(* CODESYS project PLC.project

Project tree, tasks and I/O mapping:
  Device : CODESYS Control Win V3 x64, CODESYS, version 3.5.20.40
    application Application
      libraries: Standard, 3.5.18.0 (System); MQTT Client Library, 3.5.20.1 (Stefan Roßmann Engineering Solutions)
      task MainTask (cyclic, interval t#20ms, priority 1) calls PLC_PRG, SCADA_PRG, PRG_MQTT
      Conveyers/
        function block Input_Conveyer [SFC]: free_entry, Create_Data
        function block Machine_Conveyer [SFC]: send_piece, recv_exit, Wait_entry, update_creation_state, recv_entry, rotate_exit, evaluate_entry, rotate_tool, process_exit, assemble_exit, swallow_entry
        function block Linear_Conveyor [SFC]: recv_entry
        function block Output_Conveyer [SFC]: Empty_Ramp, Reciving_entry, free_entry
        function block Unloading_Conveyer [SFC]: Extract_Data, wait_exit, clear_vars
        function block Loading_Conveyer [SFC]: load_entry
      program SCADA_PRG [ST]
      data type Piece
      program PLC_PRG [CFC]
      Symbols
      program AlarmManager [ST]
      global variables GVL
      program PRG_MQTT [ST]
      global variables GVL_MQTT
    Ethernet : Ethernet, CODESYS, version 4.2.0.0
      Modbus_TCP_Master : Modbus TCP Client, CODESYS, version 4.4.0.0
          settings: AutoReconnect = TRUE
        Modbus_TCP_Slave : Modbus TCP Server, CODESYS, version 4.4.0.0
            settings: Unit-ID = 255; IPAddress = [127, 0, 0, 1]; Port = 5502; InputChannel.Function Code = 2; InputChannel.Read Offset = 16#0000; InputChannel.Read Length = 140; InputChannel.Write Offset = 0; InputChannel.Write Length = 0; InputChannel.Cycle Time = 20; OutputChannel.Function Code = 15; OutputChannel.Read Offset = 0; OutputChannel.Read Length = 0; OutputChannel.Write Offset = 16#0000; OutputChannel.Write Length = 215; OutputChannel.Cycle Time = 20; pieces.Function Code = 16; pieces.Read Offset = 0; pieces.Read Length = 0; pieces.Write Offset = 16#0000; pieces.Write Length = 15; pieces.Cycle Time = 20
            input  Application.GVL.In[0] : BOOL  // InputChannel.InputChannel.Bit0
            input  Application.GVL.In[1] : BOOL  // InputChannel.InputChannel.Bit1
            input  Application.GVL.In[2] : BOOL  // InputChannel.InputChannel.Bit2
            input  Application.GVL.In[3] : BOOL  // InputChannel.InputChannel.Bit3
            input  Application.GVL.In[4] : BOOL  // InputChannel.InputChannel.Bit4
            input  Application.GVL.In[5] : BOOL  // InputChannel.InputChannel.Bit5
            input  Application.GVL.In[6] : BOOL  // InputChannel.InputChannel.Bit6
            input  Application.GVL.In[7] : BOOL  // InputChannel.InputChannel.Bit7
            input  Application.GVL.In[8] : BOOL  // InputChannel.InputChannel.Bit0
            input  Application.GVL.In[9] : BOOL  // InputChannel.InputChannel.Bit1
            input  Application.GVL.In[10] : BOOL  // InputChannel.InputChannel.Bit2
            input  Application.GVL.In[11] : BOOL  // InputChannel.InputChannel.Bit3
            input  Application.GVL.In[12] : BOOL  // InputChannel.InputChannel.Bit4
            input  Application.GVL.In[13] : BOOL  // InputChannel.InputChannel.Bit5
            input  Application.GVL.In[14] : BOOL  // InputChannel.InputChannel.Bit6
            input  Application.GVL.In[15] : BOOL  // InputChannel.InputChannel.Bit7
            input  Application.GVL.In[16] : BOOL  // InputChannel.InputChannel.Bit0
            input  Application.GVL.In[17] : BOOL  // InputChannel.InputChannel.Bit1
            input  Application.GVL.In[18] : BOOL  // InputChannel.InputChannel.Bit2
            input  Application.GVL.In[19] : BOOL  // InputChannel.InputChannel.Bit3
            input  Application.GVL.In[20] : BOOL  // InputChannel.InputChannel.Bit4
            input  Application.GVL.In[21] : BOOL  // InputChannel.InputChannel.Bit5
            input  Application.GVL.In[22] : BOOL  // InputChannel.InputChannel.Bit6
            input  Application.GVL.In[23] : BOOL  // InputChannel.InputChannel.Bit7
            input  Application.GVL.In[24] : BOOL  // InputChannel.InputChannel.Bit0
            input  Application.GVL.In[25] : BOOL  // InputChannel.InputChannel.Bit1
            input  Application.GVL.In[26] : BOOL  // InputChannel.InputChannel.Bit2
            input  Application.GVL.In[27] : BOOL  // InputChannel.InputChannel.Bit3
            input  Application.GVL.In[28] : BOOL  // InputChannel.InputChannel.Bit4
            input  Application.GVL.In[29] : BOOL  // InputChannel.InputChannel.Bit5
            input  Application.GVL.In[30] : BOOL  // InputChannel.InputChannel.Bit6
            input  Application.GVL.In[31] : BOOL  // InputChannel.InputChannel.Bit7
            input  Application.GVL.In[32] : BOOL  // InputChannel.InputChannel.Bit0
            input  Application.GVL.In[33] : BOOL  // InputChannel.InputChannel.Bit1
            input  Application.GVL.In[34] : BOOL  // InputChannel.InputChannel.Bit2
            input  Application.GVL.In[35] : BOOL  // InputChannel.InputChannel.Bit3
            input  Application.GVL.In[36] : BOOL  // InputChannel.InputChannel.Bit4
            input  Application.GVL.In[37] : BOOL  // InputChannel.InputChannel.Bit5
            input  Application.GVL.In[38] : BOOL  // InputChannel.InputChannel.Bit6
            input  Application.GVL.In[39] : BOOL  // InputChannel.InputChannel.Bit7
            input  Application.GVL.In[40] : BOOL  // InputChannel.InputChannel.Bit0
            input  Application.GVL.In[41] : BOOL  // InputChannel.InputChannel.Bit1
            input  Application.GVL.In[42] : BOOL  // InputChannel.InputChannel.Bit2
            input  Application.GVL.In[43] : BOOL  // InputChannel.InputChannel.Bit3
            input  Application.GVL.In[44] : BOOL  // InputChannel.InputChannel.Bit4
            input  Application.GVL.In[45] : BOOL  // InputChannel.InputChannel.Bit5
            input  Application.GVL.In[46] : BOOL  // InputChannel.InputChannel.Bit6
            input  Application.GVL.In[47] : BOOL  // InputChannel.InputChannel.Bit7
            input  Application.GVL.In[48] : BOOL  // InputChannel.InputChannel.Bit0
            input  Application.GVL.In[49] : BOOL  // InputChannel.InputChannel.Bit1
            input  Application.GVL.In[50] : BOOL  // InputChannel.InputChannel.Bit2
            input  Application.GVL.In[51] : BOOL  // InputChannel.InputChannel.Bit3
            input  Application.GVL.In[52] : BOOL  // InputChannel.InputChannel.Bit4
            input  Application.GVL.In[53] : BOOL  // InputChannel.InputChannel.Bit5
            input  Application.GVL.In[54] : BOOL  // InputChannel.InputChannel.Bit6
            input  Application.GVL.In[55] : BOOL  // InputChannel.InputChannel.Bit7
            input  Application.GVL.In[56] : BOOL  // InputChannel.InputChannel.Bit0
            input  Application.GVL.In[57] : BOOL  // InputChannel.InputChannel.Bit1
            input  Application.GVL.In[58] : BOOL  // InputChannel.InputChannel.Bit2
            input  Application.GVL.In[59] : BOOL  // InputChannel.InputChannel.Bit3
            input  Application.GVL.In[60] : BOOL  // InputChannel.InputChannel.Bit4
            input  Application.GVL.In[61] : BOOL  // InputChannel.InputChannel.Bit5
            input  Application.GVL.In[62] : BOOL  // InputChannel.InputChannel.Bit6
            input  Application.GVL.In[63] : BOOL  // InputChannel.InputChannel.Bit7
            input  Application.GVL.In[64] : BOOL  // InputChannel.InputChannel.Bit0
            input  Application.GVL.In[65] : BOOL  // InputChannel.InputChannel.Bit1
            input  Application.GVL.In[66] : BOOL  // InputChannel.InputChannel.Bit2
            input  Application.GVL.In[67] : BOOL  // InputChannel.InputChannel.Bit3
            input  Application.GVL.In[68] : BOOL  // InputChannel.InputChannel.Bit4
            input  Application.GVL.In[69] : BOOL  // InputChannel.InputChannel.Bit5
            input  Application.GVL.In[70] : BOOL  // InputChannel.InputChannel.Bit6
            input  Application.GVL.In[71] : BOOL  // InputChannel.InputChannel.Bit7
            input  Application.GVL.In[72] : BOOL  // InputChannel.InputChannel.Bit0
            input  Application.GVL.In[73] : BOOL  // InputChannel.InputChannel.Bit1
            input  Application.GVL.In[74] : BOOL  // InputChannel.InputChannel.Bit2
            input  Application.GVL.In[75] : BOOL  // InputChannel.InputChannel.Bit3
            input  Application.GVL.In[76] : BOOL  // InputChannel.InputChannel.Bit4
            input  Application.GVL.In[77] : BOOL  // InputChannel.InputChannel.Bit5
            input  Application.GVL.In[78] : BOOL  // InputChannel.InputChannel.Bit6
            input  Application.GVL.In[79] : BOOL  // InputChannel.InputChannel.Bit7
            input  Application.GVL.In[80] : BOOL  // InputChannel.InputChannel.Bit0
            input  Application.GVL.In[81] : BOOL  // InputChannel.InputChannel.Bit1
            input  Application.GVL.In[82] : BOOL  // InputChannel.InputChannel.Bit2
            input  Application.GVL.In[83] : BOOL  // InputChannel.InputChannel.Bit3
            input  Application.GVL.In[84] : BOOL  // InputChannel.InputChannel.Bit4
            input  Application.GVL.In[85] : BOOL  // InputChannel.InputChannel.Bit5
            input  Application.GVL.In[86] : BOOL  // InputChannel.InputChannel.Bit6
            input  Application.GVL.In[87] : BOOL  // InputChannel.InputChannel.Bit7
            input  Application.GVL.In[88] : BOOL  // InputChannel.InputChannel.Bit0
            input  Application.GVL.In[89] : BOOL  // InputChannel.InputChannel.Bit1
            input  Application.GVL.In[90] : BOOL  // InputChannel.InputChannel.Bit2
            input  Application.GVL.In[91] : BOOL  // InputChannel.InputChannel.Bit3
            input  Application.GVL.In[92] : BOOL  // InputChannel.InputChannel.Bit4
            input  Application.GVL.In[93] : BOOL  // InputChannel.InputChannel.Bit5
            input  Application.GVL.In[94] : BOOL  // InputChannel.InputChannel.Bit6
            input  Application.GVL.In[95] : BOOL  // InputChannel.InputChannel.Bit7
            input  Application.GVL.In[96] : BOOL  // InputChannel.InputChannel.Bit0
            input  Application.GVL.In[97] : BOOL  // InputChannel.InputChannel.Bit1
            input  Application.GVL.In[98] : BOOL  // InputChannel.InputChannel.Bit2
            input  Application.GVL.In[99] : BOOL  // InputChannel.InputChannel.Bit3
            input  Application.GVL.In[100] : BOOL  // InputChannel.InputChannel.Bit4
            input  Application.GVL.In[101] : BOOL  // InputChannel.InputChannel.Bit5
            input  Application.GVL.In[102] : BOOL  // InputChannel.InputChannel.Bit6
            input  Application.GVL.In[103] : BOOL  // InputChannel.InputChannel.Bit7
            input  Application.GVL.In[104] : BOOL  // InputChannel.InputChannel.Bit0
            input  Application.GVL.In[105] : BOOL  // InputChannel.InputChannel.Bit1
            input  Application.GVL.In[106] : BOOL  // InputChannel.InputChannel.Bit2
            input  Application.GVL.In[107] : BOOL  // InputChannel.InputChannel.Bit3
            input  Application.GVL.In[108] : BOOL  // InputChannel.InputChannel.Bit4
            input  Application.GVL.In[109] : BOOL  // InputChannel.InputChannel.Bit5
            input  Application.GVL.In[110] : BOOL  // InputChannel.InputChannel.Bit6
            input  Application.GVL.In[111] : BOOL  // InputChannel.InputChannel.Bit7
            input  Application.GVL.In[112] : BOOL  // InputChannel.InputChannel.Bit0
            input  Application.GVL.In[113] : BOOL  // InputChannel.InputChannel.Bit1
            input  Application.GVL.In[114] : BOOL  // InputChannel.InputChannel.Bit2
            input  Application.GVL.In[115] : BOOL  // InputChannel.InputChannel.Bit3
            input  Application.GVL.In[116] : BOOL  // InputChannel.InputChannel.Bit4
            input  Application.GVL.In[117] : BOOL  // InputChannel.InputChannel.Bit5
            input  Application.GVL.In[118] : BOOL  // InputChannel.InputChannel.Bit6
            input  Application.GVL.In[119] : BOOL  // InputChannel.InputChannel.Bit7
            input  Application.GVL.In[120] : BOOL  // InputChannel.InputChannel.Bit0
            input  Application.GVL.In[121] : BOOL  // InputChannel.InputChannel.Bit1
            input  Application.GVL.In[122] : BOOL  // InputChannel.InputChannel.Bit2
            input  Application.GVL.In[123] : BOOL  // InputChannel.InputChannel.Bit3
            input  Application.GVL.In[124] : BOOL  // InputChannel.InputChannel.Bit4
            input  Application.GVL.In[125] : BOOL  // InputChannel.InputChannel.Bit5
            input  Application.GVL.In[126] : BOOL  // InputChannel.InputChannel.Bit6
            input  Application.GVL.In[127] : BOOL  // InputChannel.InputChannel.Bit7
            input  Application.GVL.In[128] : BOOL  // InputChannel.InputChannel.Bit0
            input  Application.GVL.In[129] : BOOL  // InputChannel.InputChannel.Bit1
            input  Application.GVL.In[130] : BOOL  // InputChannel.InputChannel.Bit2
            input  Application.GVL.In[131] : BOOL  // InputChannel.InputChannel.Bit3
            input  Application.GVL.In[132] : BOOL  // InputChannel.InputChannel.Bit4
            input  Application.GVL.In[133] : BOOL  // InputChannel.InputChannel.Bit5
            input  Application.GVL.In[134] : BOOL  // InputChannel.InputChannel.Bit6
            input  Application.GVL.In[135] : BOOL  // InputChannel.InputChannel.Bit7
            input  Application.GVL.In[136] : BOOL  // InputChannel.InputChannel.Bit0
            input  Application.GVL.In[137] : BOOL  // InputChannel.InputChannel.Bit1
            input  Application.GVL.In[138] : BOOL  // InputChannel.InputChannel.Bit2
            input  Application.GVL.In[139] : BOOL  // InputChannel.InputChannel.Bit3
            output Application.GVL.Out[0] : BOOL  // OutputChannel.OutputChannel[0].Bit0
            output Application.GVL.Out[1] : BOOL  // OutputChannel.OutputChannel[0].Bit1
            output Application.GVL.Out[2] : BOOL  // OutputChannel.OutputChannel[0].Bit2
            output Application.GVL.Out[3] : BOOL  // OutputChannel.OutputChannel[0].Bit3
            output Application.GVL.Out[4] : BOOL  // OutputChannel.OutputChannel[0].Bit4
            output Application.GVL.Out[5] : BOOL  // OutputChannel.OutputChannel[0].Bit5
            output Application.GVL.Out[6] : BOOL  // OutputChannel.OutputChannel[0].Bit6
            output Application.GVL.Out[7] : BOOL  // OutputChannel.OutputChannel[0].Bit7
            output Application.GVL.Out[8] : BOOL  // OutputChannel.OutputChannel[1].Bit0
            output Application.GVL.Out[9] : BOOL  // OutputChannel.OutputChannel[1].Bit1
            output Application.GVL.Out[10] : BOOL  // OutputChannel.OutputChannel[1].Bit2
            output Application.GVL.Out[11] : BOOL  // OutputChannel.OutputChannel[1].Bit3
            output Application.GVL.Out[12] : BOOL  // OutputChannel.OutputChannel[1].Bit4
            output Application.GVL.Out[13] : BOOL  // OutputChannel.OutputChannel[1].Bit5
            output Application.GVL.Out[14] : BOOL  // OutputChannel.OutputChannel[1].Bit6
            output Application.GVL.Out[15] : BOOL  // OutputChannel.OutputChannel[1].Bit7
            output Application.GVL.Out[16] : BOOL  // OutputChannel.OutputChannel[2].Bit0
            output Application.GVL.Out[17] : BOOL  // OutputChannel.OutputChannel[2].Bit1
            output Application.GVL.Out[18] : BOOL  // OutputChannel.OutputChannel[2].Bit2
            output Application.GVL.Out[19] : BOOL  // OutputChannel.OutputChannel[2].Bit3
            output Application.GVL.Out[20] : BOOL  // OutputChannel.OutputChannel[2].Bit4
            output Application.GVL.Out[21] : BOOL  // OutputChannel.OutputChannel[2].Bit5
            output Application.GVL.Out[22] : BOOL  // OutputChannel.OutputChannel[2].Bit6
            output Application.GVL.Out[23] : BOOL  // OutputChannel.OutputChannel[2].Bit7
            output Application.GVL.Out[24] : BOOL  // OutputChannel.OutputChannel[3].Bit0
            output Application.GVL.Out[25] : BOOL  // OutputChannel.OutputChannel[3].Bit1
            output Application.GVL.Out[26] : BOOL  // OutputChannel.OutputChannel[3].Bit2
            output Application.GVL.Out[27] : BOOL  // OutputChannel.OutputChannel[3].Bit3
            output Application.GVL.Out[28] : BOOL  // OutputChannel.OutputChannel[3].Bit4
            output Application.GVL.Out[29] : BOOL  // OutputChannel.OutputChannel[3].Bit5
            output Application.GVL.Out[30] : BOOL  // OutputChannel.OutputChannel[3].Bit6
            output Application.GVL.Out[31] : BOOL  // OutputChannel.OutputChannel[3].Bit7
            output Application.GVL.Out[32] : BOOL  // OutputChannel.OutputChannel[4].Bit0
            output Application.GVL.Out[33] : BOOL  // OutputChannel.OutputChannel[4].Bit1
            output Application.GVL.Out[34] : BOOL  // OutputChannel.OutputChannel[4].Bit2
            output Application.GVL.Out[35] : BOOL  // OutputChannel.OutputChannel[4].Bit3
            output Application.GVL.Out[36] : BOOL  // OutputChannel.OutputChannel[4].Bit4
            output Application.GVL.Out[37] : BOOL  // OutputChannel.OutputChannel[4].Bit5
            output Application.GVL.Out[38] : BOOL  // OutputChannel.OutputChannel[4].Bit6
            output Application.GVL.Out[39] : BOOL  // OutputChannel.OutputChannel[4].Bit7
            output Application.GVL.Out[40] : BOOL  // OutputChannel.OutputChannel[5].Bit0
            output Application.GVL.Out[41] : BOOL  // OutputChannel.OutputChannel[5].Bit1
            output Application.GVL.Out[42] : BOOL  // OutputChannel.OutputChannel[5].Bit2
            output Application.GVL.Out[43] : BOOL  // OutputChannel.OutputChannel[5].Bit3
            output Application.GVL.Out[44] : BOOL  // OutputChannel.OutputChannel[5].Bit4
            output Application.GVL.Out[45] : BOOL  // OutputChannel.OutputChannel[5].Bit5
            output Application.GVL.Out[46] : BOOL  // OutputChannel.OutputChannel[5].Bit6
            output Application.GVL.Out[47] : BOOL  // OutputChannel.OutputChannel[5].Bit7
            output Application.GVL.Out[48] : BOOL  // OutputChannel.OutputChannel[6].Bit0
            output Application.GVL.Out[49] : BOOL  // OutputChannel.OutputChannel[6].Bit1
            output Application.GVL.Out[50] : BOOL  // OutputChannel.OutputChannel[6].Bit2
            output Application.GVL.Out[51] : BOOL  // OutputChannel.OutputChannel[6].Bit3
            output Application.GVL.Out[52] : BOOL  // OutputChannel.OutputChannel[6].Bit4
            output Application.GVL.Out[53] : BOOL  // OutputChannel.OutputChannel[6].Bit5
            output Application.GVL.Out[54] : BOOL  // OutputChannel.OutputChannel[6].Bit6
            output Application.GVL.Out[55] : BOOL  // OutputChannel.OutputChannel[6].Bit7
            output Application.GVL.Out[56] : BOOL  // OutputChannel.OutputChannel[7].Bit0
            output Application.GVL.Out[57] : BOOL  // OutputChannel.OutputChannel[7].Bit1
            output Application.GVL.Out[58] : BOOL  // OutputChannel.OutputChannel[7].Bit2
            output Application.GVL.Out[59] : BOOL  // OutputChannel.OutputChannel[7].Bit3
            output Application.GVL.Out[60] : BOOL  // OutputChannel.OutputChannel[7].Bit4
            output Application.GVL.Out[61] : BOOL  // OutputChannel.OutputChannel[7].Bit5
            output Application.GVL.Out[62] : BOOL  // OutputChannel.OutputChannel[7].Bit6
            output Application.GVL.Out[63] : BOOL  // OutputChannel.OutputChannel[7].Bit7
            output Application.GVL.Out[64] : BOOL  // OutputChannel.OutputChannel[8].Bit0
            output Application.GVL.Out[65] : BOOL  // OutputChannel.OutputChannel[8].Bit1
            output Application.GVL.Out[66] : BOOL  // OutputChannel.OutputChannel[8].Bit2
            output Application.GVL.Out[67] : BOOL  // OutputChannel.OutputChannel[8].Bit3
            output Application.GVL.Out[68] : BOOL  // OutputChannel.OutputChannel[8].Bit4
            output Application.GVL.Out[69] : BOOL  // OutputChannel.OutputChannel[8].Bit5
            output Application.GVL.Out[70] : BOOL  // OutputChannel.OutputChannel[8].Bit6
            output Application.GVL.Out[71] : BOOL  // OutputChannel.OutputChannel[8].Bit7
            output Application.GVL.Out[72] : BOOL  // OutputChannel.OutputChannel[9].Bit0
            output Application.GVL.Out[73] : BOOL  // OutputChannel.OutputChannel[9].Bit1
            output Application.GVL.Out[74] : BOOL  // OutputChannel.OutputChannel[9].Bit2
            output Application.GVL.Out[75] : BOOL  // OutputChannel.OutputChannel[9].Bit3
            output Application.GVL.Out[76] : BOOL  // OutputChannel.OutputChannel[9].Bit4
            output Application.GVL.Out[77] : BOOL  // OutputChannel.OutputChannel[9].Bit5
            output Application.GVL.Out[78] : BOOL  // OutputChannel.OutputChannel[9].Bit6
            output Application.GVL.Out[79] : BOOL  // OutputChannel.OutputChannel[9].Bit7
            output Application.GVL.Out[80] : BOOL  // OutputChannel.OutputChannel[10].Bit0
            output Application.GVL.Out[81] : BOOL  // OutputChannel.OutputChannel[10].Bit1
            output Application.GVL.Out[82] : BOOL  // OutputChannel.OutputChannel[10].Bit2
            output Application.GVL.Out[83] : BOOL  // OutputChannel.OutputChannel[10].Bit3
            output Application.GVL.Out[84] : BOOL  // OutputChannel.OutputChannel[10].Bit4
            output Application.GVL.Out[85] : BOOL  // OutputChannel.OutputChannel[10].Bit5
            output Application.GVL.Out[86] : BOOL  // OutputChannel.OutputChannel[10].Bit6
            output Application.GVL.Out[87] : BOOL  // OutputChannel.OutputChannel[10].Bit7
            output Application.GVL.Out[88] : BOOL  // OutputChannel.OutputChannel[11].Bit0
            output Application.GVL.Out[89] : BOOL  // OutputChannel.OutputChannel[11].Bit1
            output Application.GVL.Out[90] : BOOL  // OutputChannel.OutputChannel[11].Bit2
            output Application.GVL.Out[91] : BOOL  // OutputChannel.OutputChannel[11].Bit3
            output Application.GVL.Out[92] : BOOL  // OutputChannel.OutputChannel[11].Bit4
            output Application.GVL.Out[93] : BOOL  // OutputChannel.OutputChannel[11].Bit5
            output Application.GVL.Out[94] : BOOL  // OutputChannel.OutputChannel[11].Bit6
            output Application.GVL.Out[95] : BOOL  // OutputChannel.OutputChannel[11].Bit7
            output Application.GVL.Out[96] : BOOL  // OutputChannel.OutputChannel[12].Bit0
            output Application.GVL.Out[97] : BOOL  // OutputChannel.OutputChannel[12].Bit1
            output Application.GVL.Out[98] : BOOL  // OutputChannel.OutputChannel[12].Bit2
            output Application.GVL.Out[99] : BOOL  // OutputChannel.OutputChannel[12].Bit3
            output Application.GVL.Out[100] : BOOL  // OutputChannel.OutputChannel[12].Bit4
            output Application.GVL.Out[101] : BOOL  // OutputChannel.OutputChannel[12].Bit5
            output Application.GVL.Out[102] : BOOL  // OutputChannel.OutputChannel[12].Bit6
            output Application.GVL.Out[103] : BOOL  // OutputChannel.OutputChannel[12].Bit7
            output Application.GVL.Out[104] : BOOL  // OutputChannel.OutputChannel[13].Bit0
            output Application.GVL.Out[105] : BOOL  // OutputChannel.OutputChannel[13].Bit1
            output Application.GVL.Out[106] : BOOL  // OutputChannel.OutputChannel[13].Bit2
            output Application.GVL.Out[107] : BOOL  // OutputChannel.OutputChannel[13].Bit3
            output Application.GVL.Out[108] : BOOL  // OutputChannel.OutputChannel[13].Bit4
            output Application.GVL.Out[109] : BOOL  // OutputChannel.OutputChannel[13].Bit5
            output Application.GVL.Out[110] : BOOL  // OutputChannel.OutputChannel[13].Bit6
            output Application.GVL.Out[111] : BOOL  // OutputChannel.OutputChannel[13].Bit7
            output Application.GVL.Out[112] : BOOL  // OutputChannel.OutputChannel[14].Bit0
            output Application.GVL.Out[113] : BOOL  // OutputChannel.OutputChannel[14].Bit1
            output Application.GVL.Out[114] : BOOL  // OutputChannel.OutputChannel[14].Bit2
            output Application.GVL.Out[115] : BOOL  // OutputChannel.OutputChannel[14].Bit3
            output Application.GVL.Out[116] : BOOL  // OutputChannel.OutputChannel[14].Bit4
            output Application.GVL.Out[117] : BOOL  // OutputChannel.OutputChannel[14].Bit5
            output Application.GVL.Out[118] : BOOL  // OutputChannel.OutputChannel[14].Bit6
            output Application.GVL.Out[119] : BOOL  // OutputChannel.OutputChannel[14].Bit7
            output Application.GVL.Out[120] : BOOL  // OutputChannel.OutputChannel[15].Bit0
            output Application.GVL.Out[121] : BOOL  // OutputChannel.OutputChannel[15].Bit1
            output Application.GVL.Out[122] : BOOL  // OutputChannel.OutputChannel[15].Bit2
            output Application.GVL.Out[123] : BOOL  // OutputChannel.OutputChannel[15].Bit3
            output Application.GVL.Out[124] : BOOL  // OutputChannel.OutputChannel[15].Bit4
            output Application.GVL.Out[125] : BOOL  // OutputChannel.OutputChannel[15].Bit5
            output Application.GVL.Out[126] : BOOL  // OutputChannel.OutputChannel[15].Bit6
            output Application.GVL.Out[127] : BOOL  // OutputChannel.OutputChannel[15].Bit7
            output Application.GVL.Out[128] : BOOL  // OutputChannel.OutputChannel[16].Bit0
            output Application.GVL.Out[129] : BOOL  // OutputChannel.OutputChannel[16].Bit1
            output Application.GVL.Out[130] : BOOL  // OutputChannel.OutputChannel[16].Bit2
            output Application.GVL.Out[131] : BOOL  // OutputChannel.OutputChannel[16].Bit3
            output Application.GVL.Out[132] : BOOL  // OutputChannel.OutputChannel[16].Bit4
            output Application.GVL.Out[133] : BOOL  // OutputChannel.OutputChannel[16].Bit5
            output Application.GVL.Out[134] : BOOL  // OutputChannel.OutputChannel[16].Bit6
            output Application.GVL.Out[135] : BOOL  // OutputChannel.OutputChannel[16].Bit7
            output Application.GVL.Out[136] : BOOL  // OutputChannel.OutputChannel[17].Bit0
            output Application.GVL.Out[137] : BOOL  // OutputChannel.OutputChannel[17].Bit1
            output Application.GVL.Out[138] : BOOL  // OutputChannel.OutputChannel[17].Bit2
            output Application.GVL.Out[139] : BOOL  // OutputChannel.OutputChannel[17].Bit3
            output Application.GVL.Out[140] : BOOL  // OutputChannel.OutputChannel[17].Bit4
            output Application.GVL.Out[141] : BOOL  // OutputChannel.OutputChannel[17].Bit5
            output Application.GVL.Out[142] : BOOL  // OutputChannel.OutputChannel[17].Bit6
            output Application.GVL.Out[143] : BOOL  // OutputChannel.OutputChannel[17].Bit7
            output Application.GVL.Out[144] : BOOL  // OutputChannel.OutputChannel[18].Bit0
            output Application.GVL.Out[145] : BOOL  // OutputChannel.OutputChannel[18].Bit1
            output Application.GVL.Out[146] : BOOL  // OutputChannel.OutputChannel[18].Bit2
            output Application.GVL.Out[147] : BOOL  // OutputChannel.OutputChannel[18].Bit3
            output Application.GVL.Out[148] : BOOL  // OutputChannel.OutputChannel[18].Bit4
            output Application.GVL.Out[149] : BOOL  // OutputChannel.OutputChannel[18].Bit5
            output Application.GVL.Out[150] : BOOL  // OutputChannel.OutputChannel[18].Bit6
            output Application.GVL.Out[151] : BOOL  // OutputChannel.OutputChannel[18].Bit7
            output Application.GVL.Out[152] : BOOL  // OutputChannel.OutputChannel[19].Bit0
            output Application.GVL.Out[153] : BOOL  // OutputChannel.OutputChannel[19].Bit1
            output Application.GVL.Out[154] : BOOL  // OutputChannel.OutputChannel[19].Bit2
            output Application.GVL.Out[155] : BOOL  // OutputChannel.OutputChannel[19].Bit3
            output Application.GVL.Out[156] : BOOL  // OutputChannel.OutputChannel[19].Bit4
            output Application.GVL.Out[157] : BOOL  // OutputChannel.OutputChannel[19].Bit5
            output Application.GVL.Out[158] : BOOL  // OutputChannel.OutputChannel[19].Bit6
            output Application.GVL.Out[159] : BOOL  // OutputChannel.OutputChannel[19].Bit7
            output Application.GVL.Out[160] : BOOL  // OutputChannel.OutputChannel[20].Bit0
            output Application.GVL.Out[161] : BOOL  // OutputChannel.OutputChannel[20].Bit1
            output Application.GVL.Out[162] : BOOL  // OutputChannel.OutputChannel[20].Bit2
            output Application.GVL.Out[163] : BOOL  // OutputChannel.OutputChannel[20].Bit3
            output Application.GVL.Out[164] : BOOL  // OutputChannel.OutputChannel[20].Bit4
            output Application.GVL.Out[165] : BOOL  // OutputChannel.OutputChannel[20].Bit5
            output Application.GVL.Out[166] : BOOL  // OutputChannel.OutputChannel[20].Bit6
            output Application.GVL.Out[167] : BOOL  // OutputChannel.OutputChannel[20].Bit7
            output Application.GVL.Out[168] : BOOL  // OutputChannel.OutputChannel[21].Bit0
            output Application.GVL.Out[169] : BOOL  // OutputChannel.OutputChannel[21].Bit1
            output Application.GVL.Out[170] : BOOL  // OutputChannel.OutputChannel[21].Bit2
            output Application.GVL.Out[171] : BOOL  // OutputChannel.OutputChannel[21].Bit3
            output Application.GVL.Out[172] : BOOL  // OutputChannel.OutputChannel[21].Bit4
            output Application.GVL.Out[173] : BOOL  // OutputChannel.OutputChannel[21].Bit5
            output Application.GVL.Out[174] : BOOL  // OutputChannel.OutputChannel[21].Bit6
            output Application.GVL.Out[175] : BOOL  // OutputChannel.OutputChannel[21].Bit7
            output Application.GVL.Out[176] : BOOL  // OutputChannel.OutputChannel[22].Bit0
            output Application.GVL.Out[177] : BOOL  // OutputChannel.OutputChannel[22].Bit1
            output Application.GVL.Out[178] : BOOL  // OutputChannel.OutputChannel[22].Bit2
            output Application.GVL.Out[179] : BOOL  // OutputChannel.OutputChannel[22].Bit3
            output Application.GVL.Out[180] : BOOL  // OutputChannel.OutputChannel[22].Bit4
            output Application.GVL.Out[181] : BOOL  // OutputChannel.OutputChannel[22].Bit5
            output Application.GVL.Out[182] : BOOL  // OutputChannel.OutputChannel[22].Bit6
            output Application.GVL.Out[183] : BOOL  // OutputChannel.OutputChannel[22].Bit7
            output Application.GVL.Out[184] : BOOL  // OutputChannel.OutputChannel[23].Bit0
            output Application.GVL.Out[185] : BOOL  // OutputChannel.OutputChannel[23].Bit1
            output Application.GVL.Out[186] : BOOL  // OutputChannel.OutputChannel[23].Bit2
            output Application.GVL.Out[187] : BOOL  // OutputChannel.OutputChannel[23].Bit3
            output Application.GVL.Out[188] : BOOL  // OutputChannel.OutputChannel[23].Bit4
            output Application.GVL.Out[189] : BOOL  // OutputChannel.OutputChannel[23].Bit5
            output Application.GVL.Out[190] : BOOL  // OutputChannel.OutputChannel[23].Bit6
            output Application.GVL.Out[191] : BOOL  // OutputChannel.OutputChannel[23].Bit7
            output Application.GVL.Out[192] : BOOL  // OutputChannel.OutputChannel[24].Bit0
            output Application.GVL.Out[193] : BOOL  // OutputChannel.OutputChannel[24].Bit1
            output Application.GVL.Out[194] : BOOL  // OutputChannel.OutputChannel[24].Bit2
            output Application.GVL.Out[195] : BOOL  // OutputChannel.OutputChannel[24].Bit3
            output Application.GVL.Out[196] : BOOL  // OutputChannel.OutputChannel[24].Bit4
            output Application.GVL.Out[197] : BOOL  // OutputChannel.OutputChannel[24].Bit5
            output Application.GVL.Out[198] : BOOL  // OutputChannel.OutputChannel[24].Bit6
            output Application.GVL.Out[199] : BOOL  // OutputChannel.OutputChannel[24].Bit7
            output Application.GVL.Out[200] : BOOL  // OutputChannel.OutputChannel[25].Bit0
            output Application.GVL.Out[201] : BOOL  // OutputChannel.OutputChannel[25].Bit1
            output Application.GVL.Out[202] : BOOL  // OutputChannel.OutputChannel[25].Bit2
            output Application.GVL.Out[203] : BOOL  // OutputChannel.OutputChannel[25].Bit3
            output Application.GVL.Out[204] : BOOL  // OutputChannel.OutputChannel[25].Bit4
            output Application.GVL.Out[205] : BOOL  // OutputChannel.OutputChannel[25].Bit5
            output Application.GVL.Out[206] : BOOL  // OutputChannel.OutputChannel[25].Bit6
            output Application.GVL.Out[207] : BOOL  // OutputChannel.OutputChannel[25].Bit7
            output Application.GVL.Out[208] : BOOL  // OutputChannel.OutputChannel[26].Bit0
            output Application.GVL.Out[209] : BOOL  // OutputChannel.OutputChannel[26].Bit1
            output Application.GVL.Out[210] : BOOL  // OutputChannel.OutputChannel[26].Bit2
            output Application.GVL.Out[211] : BOOL  // OutputChannel.OutputChannel[26].Bit3
            output Application.GVL.Out[212] : BOOL  // OutputChannel.OutputChannel[26].Bit4
            output Application.GVL.Out[213] : BOOL  // OutputChannel.OutputChannel[26].Bit5
            output Application.GVL.Out[214] : BOOL  // OutputChannel.OutputChannel[26].Bit6
            output Application.GVL.Reg[0] : WORD  // pieces.pieces[0]
            output Application.GVL.Reg[1] : WORD  // pieces.pieces[1]
            output Application.GVL.Reg[2] : WORD  // pieces.pieces[2]
            output Application.GVL.Reg[3] : WORD  // pieces.pieces[3]
            output Application.GVL.Reg[4] : WORD  // pieces.pieces[4]
            output Application.GVL.Reg[5] : WORD  // pieces.pieces[5]
            output Application.GVL.Reg[6] : WORD  // pieces.pieces[6]
            output Application.GVL.Reg[7] : WORD  // pieces.pieces[7]
            output Application.GVL.Reg[8] : WORD  // pieces.pieces[8]
            output Application.GVL.Reg[9] : WORD  // pieces.pieces[9]
            output Application.GVL.Reg[10] : WORD  // pieces.pieces[10]
            output Application.GVL.Reg[11] : WORD  // pieces.pieces[11]
            output Application.GVL.Reg[12] : WORD  // pieces.pieces[12]
            output Application.GVL.Reg[13] : WORD  // pieces.pieces[13]
            output Application.GVL.Reg[14] : WORD  // pieces.pieces[14]
            unmapped channels: InputChannel, OutputChannel, pieces
      ModbusTCP_Slave_Device : ModbusTCP Server Device, CODESYS, version 4.4.0.0
          settings: UpdateableHolding = TRUE; DistinctBitAreas = TRUE; Coils Size = 48; Discrete Inputs Size = 8
          output S_sensor1 : BOOL  // Holding Registers.Holding Registers.Bit0
          output S_sensor2 : BOOL  // Holding Registers.Holding Registers.Bit1
          output S_sensor3 : BOOL  // Holding Registers.Holding Registers.Bit2
          output C1_stop : BOOL  // Holding Registers.Holding Registers.Bit0
          output C2_stop : BOOL  // Holding Registers.Holding Registers.Bit1
          output C3_stop : BOOL  // Holding Registers.Holding Registers.Bit2
          output In_on : BOOL  // Coils.Coils.Bit0
          output M1a_on : BOOL  // Coils.Coils.Bit1
          output L1_on : BOOL  // Coils.Coils.Bit2
          output M1b_on : BOOL  // Coils.Coils.Bit3
          output L2_on : BOOL  // Coils.Coils.Bit4
          output M1c_on : BOOL  // Coils.Coils.Bit5
          output Out_on : BOOL  // Coils.Coils.Bit6
          output C1_In_Sensor : BOOL  // Coils.Coils.Bit7
          output M1a_Sensor : BOOL  // Coils.Coils.Bit0
          output C1_L1_Sensor : BOOL  // Coils.Coils.Bit1
          output M1b_Sensor : BOOL  // Coils.Coils.Bit2
          output C1_L2_Sensor : BOOL  // Coils.Coils.Bit3
          output M1c_Sensor : BOOL  // Coils.Coils.Bit4
          output M1a_T1 : BOOL  // Coils.Coils.Bit5
          output M1a_T2 : BOOL  // Coils.Coils.Bit6
          output M1a_T3 : BOOL  // Coils.Coils.Bit7
          output C1_Out_Sensor : BOOL  // Coils.Coils.Bit0
          output M1a_done : BOOL  // Coils.Coils.Bit1
          output M1a_Idle_Alarm : BOOL  // Coils.Coils.Bit2
          output M1a_Manual : BOOL  // Coils.Coils.Bit3
          output M1a_Auto : BOOL  // Coils.Coils.Bit4
          output M1c_T11 : BOOL  // Coils.Coils.Bit5
          output M1a_Manutencao : BOOL  // Coils.Coils.Bit6
          unmapped channels: Holding Registers, Input Registers, Coils, Discrete Inputs
*)

// Device/Application/Piece
TYPE Piece :
STRUCT
	/// 0=Empty, 1=Wood, 2=Metal, 3=RtopW, 4=STopW, 5=LegW, 6=RtopM, 7=STopM, 8=LegM, 9=RWW, 10=SWW, 11=RWM, 12=SWM, 13=RMM, 14=SMM
	Type_ID: UINT;
	/// TRUE if piece is destroyed 
	Is_Black: BOOL;
END_STRUCT
END_TYPE

// Device/Application/GVL
VAR_GLOBAL
	In: ARRAY[0..139] OF BOOL;
	Out: ARRAY[0..220] OF BOOL;
	Reg: ARRAY[0..15] OF UINT;
	WareHouseTop: ARRAY[0..31] OF Piece;
	WareHouseBottom: ARRAY[0..31] OF Piece;
	/// Number of pieces currently in W1
	W1_Count: UINT := 0;
	/// Number of pieces currently in W2~
	W2_Count: UINT := 0;
	
	Tool_M1a: ARRAY[0..2] OF INT := [1, 2, 3];
	Tool_Time: ARRAY[0..11] OF TIME := [T#0S, T#30S, T#20S, T#10S, T#35S, T#30S, T#25S, T#0S, T#10S, T#10S, T#30S, T#40S];
	Tool_M1b: ARRAY[0..2] OF INT := [1, 2, 3];
	Tool_M1c: ARRAY[0..2] OF INT := [8, 9, 11];
	Tool_M2a: ARRAY[0..2] OF INT := [1, 2, 3];
	Tool_M2b: ARRAY[0..2] OF INT := [1, 2, 3];
	Tool_M2c: ARRAY[0..2] OF INT := [8, 9, 10];
	Tool_M3a: ARRAY[0..2] OF INT := [4, 5, 6];
	Tool_M3b: ARRAY[0..2] OF INT := [4, 5, 6];
	Tool_M3c: ARRAY[0..2] OF INT := [8, 9, 11];
	Tool_M4a: ARRAY[0..2] OF INT := [4, 5, 6];
	Tool_M4b: ARRAY[0..2] OF INT := [4, 5, 6];
	Tool_M4c: ARRAY[0..2] OF INT := [8, 9, 10];
END_VAR

// Device/Application/GVL_MQTT
(*
  GVL_MQTT — Global Variable List for ThingsBoard MQTT connection
  Paste this into a new GVL named "GVL_MQTT" in CODESYS.
  Requires: MQTT Client Library (namespace: MQTT_Client) in Library Manager.
*)

VAR_GLOBAL
    // Publisher — sends PLC I/O telemetry to ThingsBoard PLC_Gateway device
    fbMQTT_Pub          : MQTT_Client.FB_MQTTClient;

    // Subscriber — receives RPC commands from ThingsBoard
    fbMQTT_Sub          : MQTT_Client.FB_MQTTClient;

    // 2-second publish timer
    tPublishTimer       : TON;

    // Publish group counter (1=inputs, 2=unload req, 3=unload type, 4=warehouse)
    nPublishGroup       : INT := 0;

    // RPC command handling
    sRPCMessage         : STRING(1024);
    bNewRPC             : BOOL;
	
END_VAR

// Device/Application/PLC_PRG
PROGRAM PLC_PRG
VAR
	C1: Linear_Conveyor;
	C2: Linear_Conveyor;
	C3: Linear_Conveyor;
	C4: Linear_Conveyor;
	C5: Linear_Conveyor;
	C7: Linear_Conveyor;
	C9: Linear_Conveyor;
	C12: Linear_Conveyor;
	C14: Linear_Conveyor;
	C17: Linear_Conveyor;
	C19: Linear_Conveyor;
	C22: Linear_Conveyor;
	C24: Linear_Conveyor;
	C6: Machine_Conveyer;
	C8: Machine_Conveyer;
	C10: Machine_Conveyer;
	C11: Machine_Conveyer;
	C13: Machine_Conveyer;
	C15: Machine_Conveyer;
	C16: Machine_Conveyer;
	C18: Machine_Conveyer;
	C20: Machine_Conveyer;
	C21: Machine_Conveyer;
	C23: Machine_Conveyer;
	C25: Machine_Conveyer;
	O1: Output_Conveyer;
	O2: Output_Conveyer;
	O3: Output_Conveyer;
	O4: Output_Conveyer;
	O5: Output_Conveyer;
	I1: Input_Conveyer;
	I2: Input_Conveyer;
	I3: Input_Conveyer;
	I4: Input_Conveyer;
	I5: Input_Conveyer;
	U1: Unloading_Conveyer;
	U2: Unloading_Conveyer;
	U3: Unloading_Conveyer;
	U4: Unloading_Conveyer;
	U5: Unloading_Conveyer;
	U6: Unloading_Conveyer;
	U7: Unloading_Conveyer;
	U8: Unloading_Conveyer;
	U9: Unloading_Conveyer;
	U10: Unloading_Conveyer;
	L1: Loading_Conveyer;
	L2: Loading_Conveyer;
	L3: Loading_Conveyer;
	L4: Loading_Conveyer;
	L5: Loading_Conveyer;
	L6: Loading_Conveyer;
	L7: Loading_Conveyer;
	L8: Loading_Conveyer;
	L9: Loading_Conveyer;
	L10: Loading_Conveyer;
	piece_material_I1: UINT;
	piece_material_I2: UINT;
	piece_material_I3: UINT;
	piece_material_I4: UINT;
	piece_material_I5: UINT;
	piece_material_U1: UINT;
	piece_material_U2: UINT;
	piece_material_U3: UINT;
	piece_material_U4: UINT;
	piece_material_U5: UINT;
	piece_material_U6: UINT;
	piece_material_U7: UINT;
	piece_material_U8: UINT;
	piece_material_U9: UINT;
	piece_material_U10: UINT;
	Create_Piece_I1: BOOL;
	Create_Piece_I2: BOOL;
	Create_Piece_I3: BOOL;
	Create_Piece_I4: BOOL;
	Create_Piece_I5: BOOL;
	Unload_Req_U1: BOOL;
	Unload_Req_U2: BOOL;
	Unload_Req_U3: BOOL;
	Unload_Req_U4: BOOL;
	Unload_Req_U5: BOOL;
	Unload_Req_U6: BOOL;
	Unload_Req_U7: BOOL;
	Unload_Req_U8: BOOL;
	Unload_Req_U9: BOOL;
	Unload_Req_U10: BOOL;
	Unload_Type_U1: UINT;
	Unload_Type_U2: UINT;
	Unload_Type_U3: UINT;
	Unload_Type_U4: UINT;
	Unload_Type_U5: UINT;
	Unload_Type_U6: UINT;
	Unload_Type_U7: UINT;
	Unload_Type_U8: UINT;
	Unload_Type_U9: UINT;
	Unload_Type_U10: UINT;
	Output_Unload_O1: BOOL;
	Output_Unload_O2: BOOL;
	Output_Unload_O3: BOOL;
	Output_Unload_O4: BOOL;
	Output_Unload_O5: BOOL;
END_VAR

I1(
    Ioff := 0,
    Qoff := 0,
    Create_Piece := Create_Piece_I1,
    piece_material := piece_material_I1,
    free_I := L6.free_O,
    reg_numb := 0); // Input_Conveyer
L6(Ioff := 5, Qoff := 10, Target_WH := 1, Direction := 1, Piece_In := I1.Piece_Out, recv_I := I1.recv_O); // Loading_Conveyer
I2(
    Ioff := 1,
    Qoff := 2,
    Create_Piece := Create_Piece_I2,
    piece_material := piece_material_I2,
    free_I := L7.free_O,
    reg_numb := 1); // Input_Conveyer
L7(Ioff := 6, Qoff := 13, Target_WH := 1, Direction := 1, Piece_In := I2.Piece_Out, recv_I := I2.recv_O); // Loading_Conveyer
I3(
    Ioff := 2,
    Qoff := 4,
    Create_Piece := Create_Piece_I3,
    piece_material := piece_material_I3,
    free_I := L8.free_O,
    reg_numb := 2); // Input_Conveyer
L8(Ioff := 7, Qoff := 16, Target_WH := 1, Direction := 1, Piece_In := I3.Piece_Out, recv_I := I3.recv_O); // Loading_Conveyer
I4(
    Ioff := 3,
    Qoff := 6,
    Create_Piece := Create_Piece_I4,
    piece_material := piece_material_I4,
    free_I := L9.free_O,
    reg_numb := 3); // Input_Conveyer
L9(Ioff := 8, Qoff := 19, Target_WH := 1, Direction := 1, Piece_In := I4.Piece_Out, recv_I := I4.recv_O); // Loading_Conveyer
I5(
    Ioff := 4,
    Qoff := 8,
    Create_Piece := Create_Piece_I5,
    piece_material := piece_material_I5,
    free_I := L10.free_O,
    reg_numb := 4); // Input_Conveyer
L10(Ioff := 9, Qoff := 22, Target_WH := 1, Direction := 1, Piece_In := I5.Piece_Out, recv_I := I5.recv_O); // Loading_Conveyer
L1(Ioff := 10, Qoff := 25, Target_WH := 1, Direction := 0, Piece_In := C1.Passed_Piece, recv_I := C1.recv_O); // Loading_Conveyer
U2(
    Ioff := 11,
    Qoff := 28,
    Target_WH := 1,
    Direction := 1,
    Unload_Req := Unload_Req_U2,
    free_I := C6.free_O,
    piece_material := Unload_Type_U2,
    reg_numb := 5); // Unloading_Conveyer
U3(
    Ioff := 12,
    Qoff := 30,
    Target_WH := 1,
    Direction := 1,
    Unload_Req := Unload_Req_U3,
    free_I := C11.free_O,
    piece_material := Unload_Type_U3,
    reg_numb := 6); // Unloading_Conveyer
U4(
    Ioff := 13,
    Qoff := 32,
    Target_WH := 1,
    Direction := 1,
    Unload_Req := Unload_Req_U4,
    free_I := C16.free_O,
    piece_material := Unload_Type_U4,
    reg_numb := 7); // Unloading_Conveyer
U5(
    Ioff := 14,
    Qoff := 34,
    Target_WH := 1,
    Direction := 1,
    Unload_Req := Unload_Req_U5,
    free_I := C21.free_O,
    piece_material := Unload_Type_U5,
    reg_numb := 8); // Unloading_Conveyer
C1(
    Ioff := 25,
    Qoff := 60,
    Direction := 0,
    Piece_Type := C2.Passed_Piece,
    recv_I := C2.recv_O,
    free_I := L1.free_O); // Linear_Conveyor
C6(
    Ioff := 30,
    Qoff := 70,
    Piece_In := U2.Piece_Out,
    recv_I := U2.recv_O,
    Direction := 1,
    free_I := C7.free_O,
    Tool_Magazine := GVL.Tool_M1a); // Machine_Conveyer
C11(
    Ioff := 50,
    Qoff := 104,
    Piece_In := U3.Piece_Out,
    recv_I := U3.recv_O,
    Direction := 1,
    free_I := C12.free_O,
    Tool_Magazine := GVL.Tool_M2a); // Machine_Conveyer
C16(
    Ioff := 70,
    Qoff := 138,
    Piece_In := U4.Piece_Out,
    recv_I := U4.recv_O,
    Direction := 1,
    free_I := C17.free_O,
    Tool_Magazine := GVL.Tool_M3a); // Machine_Conveyer
C21(
    Ioff := 90,
    Qoff := 172,
    Piece_In := U5.Piece_Out,
    Direction := 1,
    recv_I := U5.recv_O,
    free_I := C22.free_O,
    Tool_Magazine := GVL.Tool_M4a); // Machine_Conveyer
C2(
    Ioff := 26,
    Qoff := 62,
    Direction := 0,
    Piece_Type := C3.Passed_Piece,
    recv_I := C3.recv_O,
    free_I := C1.free_O); // Linear_Conveyor
C7(
    Ioff := 36,
    Qoff := 80,
    Direction := 1,
    Piece_Type := C6.Piece_Out,
    recv_I := C6.recv_O,
    free_I := C8.free_O); // Linear_Conveyor
C12(
    Ioff := 56,
    Qoff := 114,
    Direction := 1,
    Piece_Type := C11.Piece_Out,
    recv_I := C11.recv_O,
    free_I := C13.free_O); // Linear_Conveyor
C17(
    Ioff := 76,
    Qoff := 148,
    Direction := 1,
    Piece_Type := C16.Piece_Out,
    recv_I := C16.recv_O,
    free_I := C18.free_O); // Linear_Conveyor
C22(
    Ioff := 96,
    Qoff := 182,
    Direction := 1,
    Piece_Type := C21.Piece_Out,
    recv_I := C21.recv_O,
    free_I := C23.free_O); // Linear_Conveyor
C3(
    Ioff := 27,
    Qoff := 64,
    Direction := 0,
    Piece_Type := C4.Passed_Piece,
    recv_I := C4.recv_O,
    free_I := C2.free_O); // Linear_Conveyor
C8(
    Ioff := 37,
    Qoff := 82,
    Piece_In := C7.Passed_Piece,
    Direction := 1,
    recv_I := C7.recv_O,
    free_I := C9.free_O,
    Tool_Magazine := GVL.Tool_M1b); // Machine_Conveyer
C13(
    Ioff := 57,
    Qoff := 116,
    Piece_In := C12.Passed_Piece,
    Direction := 1,
    recv_I := C12.recv_O,
    free_I := C14.free_O,
    Tool_Magazine := GVL.Tool_M2b); // Machine_Conveyer
C18(
    Ioff := 77,
    Qoff := 150,
    Piece_In := C17.Passed_Piece,
    Direction := 1,
    recv_I := C17.recv_O,
    free_I := C19.free_O,
    Tool_Magazine := GVL.Tool_M3b); // Machine_Conveyer
C23(
    Ioff := 97,
    Qoff := 184,
    Piece_In := C22.Passed_Piece,
    Direction := 1,
    recv_I := C22.recv_O,
    free_I := C24.free_O,
    Tool_Magazine := GVL.Tool_M4b); // Machine_Conveyer
C4(
    Ioff := 28,
    Qoff := 66,
    Direction := 0,
    Piece_Type := C5.Passed_Piece,
    recv_I := C5.recv_O,
    free_I := C3.free_O); // Linear_Conveyor
C9(
    Ioff := 43,
    Qoff := 92,
    Direction := 1,
    Piece_Type := C8.Piece_Out,
    recv_I := C8.recv_O,
    free_I := C10.free_O); // Linear_Conveyor
C14(
    Ioff := 63,
    Qoff := 126,
    Direction := 1,
    Piece_Type := C13.Piece_Out,
    recv_I := C13.recv_O,
    free_I := C15.free_O); // Linear_Conveyor
C19(
    Ioff := 83,
    Qoff := 160,
    Direction := 1,
    Piece_Type := C18.Piece_Out,
    recv_I := C18.recv_O,
    free_I := C20.free_O); // Linear_Conveyor
C24(
    Ioff := 103,
    Qoff := 194,
    Direction := 1,
    Piece_Type := C23.Piece_Out,
    recv_I := C23.recv_O,
    free_I := C25.free_O); // Linear_Conveyor
C5(
    Ioff := 29,
    Qoff := 68,
    Direction := 0,
    Piece_Type := U1.Piece_Out,
    recv_I := U1.recv_O,
    free_I := C4.free_O); // Linear_Conveyor
U1(
    Ioff := 20,
    Qoff := 46,
    Target_WH := 2,
    Direction := 0,
    Unload_Req := Unload_Req_U1,
    free_I := C5.free_O,
    piece_material := Unload_Type_U1,
    reg_numb := 14); // Unloading_Conveyer
C10(
    Ioff := 44,
    Qoff := 94,
    Piece_In := C9.Passed_Piece,
    Direction := 1,
    recv_I := C9.recv_O,
    free_I := L2.free_O,
    Tool_Magazine := GVL.Tool_M1c); // Machine_Conveyer
L2(Ioff := 21, Qoff := 48, Target_WH := 2, Direction := 1, Piece_In := C10.Piece_Out, recv_I := C10.recv_O); // Loading_Conveyer
C15(
    Ioff := 64,
    Qoff := 128,
    Piece_In := C14.Passed_Piece,
    Direction := 1,
    recv_I := C14.recv_O,
    free_I := L3.free_O,
    Tool_Magazine := GVL.Tool_M2c); // Machine_Conveyer
L3(Ioff := 22, Qoff := 51, Target_WH := 2, Direction := 1, Piece_In := C15.Piece_Out, recv_I := C15.recv_O); // Loading_Conveyer
C20(
    Ioff := 84,
    Qoff := 162,
    Piece_In := C19.Passed_Piece,
    Direction := 1,
    recv_I := C19.recv_O,
    free_I := L4.free_O,
    Tool_Magazine := GVL.Tool_M3c); // Machine_Conveyer
L4(Ioff := 23, Qoff := 54, Target_WH := 2, Direction := 1, Piece_In := C20.Piece_Out, recv_I := C20.recv_O); // Loading_Conveyer
C25(
    Ioff := 104,
    Qoff := 196,
    Piece_In := C24.Passed_Piece,
    Direction := 1,
    recv_I := C24.recv_O,
    free_I := L5.free_O,
    Tool_Magazine := GVL.Tool_M4c); // Machine_Conveyer
L5(Ioff := 24, Qoff := 57, Target_WH := 2, Direction := 1, Piece_In := C25.Piece_Out, recv_I := C25.recv_O); // Loading_Conveyer
U6(
    Ioff := 15,
    Qoff := 36,
    Target_WH := 2,
    Direction := 1,
    Unload_Req := Unload_Req_U6,
    free_I := O1.free_O,
    piece_material := Unload_Type_U6,
    reg_numb := 9); // Unloading_Conveyer
O1(Ioff := 110, Qoff := 206, recv_I := U6.recv_O, Piece_In := U6.Piece_Out, Unload_Cmd := Output_Unload_O1); // Output_Conveyer
U7(
    Ioff := 16,
    Qoff := 38,
    Target_WH := 2,
    Direction := 1,
    Unload_Req := Unload_Req_U7,
    free_I := O2.free_O,
    piece_material := Unload_Type_U7,
    reg_numb := 10); // Unloading_Conveyer
O2(Ioff := 116, Qoff := 208, recv_I := U7.recv_O, Piece_In := U7.Piece_Out, Unload_Cmd := Output_Unload_O2); // Output_Conveyer
U8(
    Ioff := 17,
    Qoff := 40,
    Target_WH := 2,
    Direction := 1,
    Unload_Req := Unload_Req_U8,
    free_I := O3.free_O,
    piece_material := Unload_Type_U8,
    reg_numb := 11); // Unloading_Conveyer
O3(Ioff := 122, Qoff := 210, recv_I := U8.recv_O, Piece_In := U8.Piece_Out, Unload_Cmd := Output_Unload_O3); // Output_Conveyer
U9(
    Ioff := 18,
    Qoff := 42,
    Target_WH := 2,
    Direction := 1,
    Unload_Req := Unload_Req_U9,
    free_I := O4.free_O,
    piece_material := Unload_Type_U9,
    reg_numb := 12); // Unloading_Conveyer
O4(Ioff := 128, Qoff := 212, recv_I := U9.recv_O, Piece_In := U9.Piece_Out, Unload_Cmd := Output_Unload_O4); // Output_Conveyer
U10(
    Ioff := 19,
    Qoff := 44,
    Target_WH := 2,
    Direction := 1,
    Unload_Req := Unload_Req_U10,
    free_I := O5.free_O,
    piece_material := Unload_Type_U10,
    reg_numb := 13); // Unloading_Conveyer
O5(Ioff := 134, Qoff := 214, recv_I := U10.recv_O, Piece_In := U10.Piece_Out, Unload_Cmd := Output_Unload_O5); // Output_Conveyer

END_PROGRAM

// Device/Application/Conveyers/Output_Conveyer
{attribute 'do_checks_for_implicit_code' := ''}
FUNCTION_BLOCK Output_Conveyer
VAR_OUTPUT
	/// TRUE when belt is empty
	free_O: BOOL;
END_VAR
VAR_INPUT
	/// Modbus index for the FIRST sensor 
	Ioff: INT;
	/// Modbus index for the FIRST motor 
	Qoff: INT;
	/// TRUE when previus belt wants to send a piece
	recv_I: BOOL;
	Piece_In: Piece;
	/// Command to flush the ramp
	Unload_Cmd: BOOL;
END_VAR
VAR
	EMPTY: BOOL;
	Has_Piece: BOOL := FALSE;
	Piece_Count: INT;
	i: INT;
	O_Unload_Timer : TON;
END_VAR

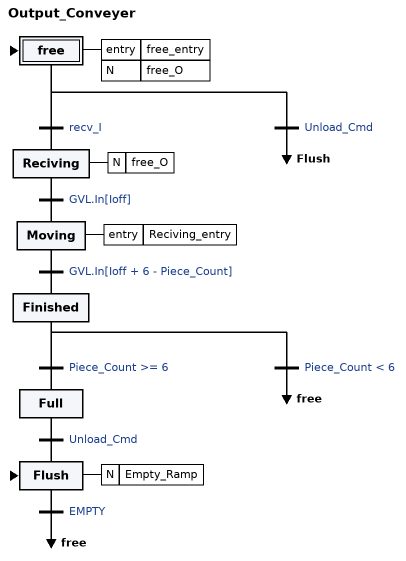
INITIAL_STEP free:
    free_entry(P1);  // entry action
    free_O(N);
END_STEP
TRANSITION FROM free TO Reciving
    := recv_I;
END_TRANSITION
STEP Reciving:
    free_O(N);
END_STEP
TRANSITION FROM Reciving TO Moving
    := GVL.In[Ioff];
END_TRANSITION
TRANSITION FROM free TO Flush
    := Unload_Cmd;
END_TRANSITION
STEP Moving:
    Reciving_entry(P1);  // entry action
END_STEP
TRANSITION FROM Moving TO Finished
    := GVL.In[Ioff + 6 - Piece_Count];
END_TRANSITION
STEP Finished:
END_STEP
TRANSITION FROM Finished TO Full
    := Piece_Count >= 6;
END_TRANSITION
STEP Full:
END_STEP
TRANSITION FROM Full TO Flush
    := Unload_Cmd;
END_TRANSITION
TRANSITION FROM Finished TO free
    := Piece_Count < 6;
END_TRANSITION
STEP Flush:
    Empty_Ramp(N);
END_STEP
TRANSITION FROM Flush TO free
    := EMPTY;
END_TRANSITION

ACTION Empty_Ramp:

Has_Piece := FALSE;
FOR i := 0 TO 6 DO
	IF(GVL.In[Ioff + 6 - i] = TRUE) THEN
		Has_Piece := TRUE;
	END_IF
END_FOR


GVL.Out[Qoff + 1] := TRUE; 


IF NOT Has_Piece THEN
	GVL.Out[Qoff + 1] := FALSE;
	EMPTY := TRUE;
	Piece_Count := 0;
END_IF




// IF (GVL.In[Ioff + 5]) AND Has_Piece THEN
// 	Piece_Count := Piece_count - 1;
// ELSE
// 	Has_Piece := TRUE;
// END_IF
// 
// IF NOT (GVL.In[Ioff + 5]) THEN
// 	Has_Piece := FALSE;
// END_IF
// 
// IF Piece_Count >= 0 THEN
// 	GVL.Out[Qoff + 1] := TRUE; 
// ELSE
// 	GVL.Out[Qoff + 1] := FALSE;
// 	EMPTY := TRUE;
// 	Piece_Count := 0;
// END_IF

// O_Unload_Timer(IN := TRUE, PT := T#6S);
// 
// IF O_Unload_Timer.Q THEN
//     EMPTY := TRUE;       // auto-close after 5s
// 	Piece_Count := 0;
//     O_Unload_Timer(IN := FALSE);    // reset timer
// END_IF
END_ACTION

ACTION Reciving_entry:
Piece_Count := Piece_Count + 1;
END_ACTION

ACTION free_entry:
EMPTY := FALSE;
END_ACTION

END_FUNCTION_BLOCK

// Device/Application/Conveyers/Loading_Conveyer
{attribute 'do_checks_for_implicit_code' := ''}
FUNCTION_BLOCK Loading_Conveyer
VAR_OUTPUT
	/// TRUE when belt is empty
	free_O: BOOL;
END_VAR
VAR
	/// Iterator for the FOR loop
	i: INT;
	/// Internal flag
	Stored: BOOL;
END_VAR
VAR_INPUT
	/// Modbus index for the sensor
	Ioff: UINT;
	/// Modbus index for the motor
	Qoff: UINT;
	/// 1 = Top (W1), 2 = Bottom (W2)
	Target_WH: INT;
	/// 0 for going UP , 1 for going DOWN
	Direction: UINT;
	/// Code for the piece 
	Piece_In: Piece;
	/// TRUE when previus belt wants to send a piece
	recv_I: BOOL;
END_VAR

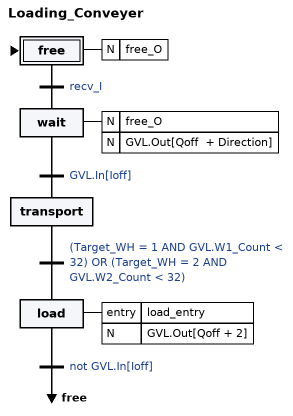
INITIAL_STEP free:
    free_O(N);
END_STEP
TRANSITION FROM free TO wait
    := recv_I;
END_TRANSITION
STEP wait:
    free_O(N);
    GVL.Out[Qoff  + Direction](N);
END_STEP
TRANSITION FROM wait TO transport
    := GVL.In[Ioff];
END_TRANSITION
STEP transport:
END_STEP
TRANSITION FROM transport TO load
    := (Target_WH = 1 AND GVL.W1_Count < 32) OR (Target_WH = 2 AND GVL.W2_Count < 32);
END_TRANSITION
STEP load:
    load_entry(P1);  // entry action
    GVL.Out[Qoff + 2](N);
END_STEP
TRANSITION FROM load TO free
    := not GVL.In[Ioff];
END_TRANSITION

ACTION load_entry:
IF Target_WH = 1 THEN
	// Save the incoming piece data into the array
	GVL.WareHouseTop[GVL.W1_Count] := Piece_In;
	
	// Update the SCADA counter
	GVL.W1_Count := GVL.W1_Count + 1;
	
// --- TARGETING BOTTOM WAREHOUSE (W2) ---
ELSIF Target_WH = 2 THEN

	// Save the incoming piece data into the array
	GVL.WareHouseBottom[GVL.W2_Count] := Piece_In;
	
	// Update the SCADA counter
	GVL.W2_Count := GVL.W2_Count + 1;

END_IF;
END_ACTION

END_FUNCTION_BLOCK

// Device/Application/Conveyers/Unloading_Conveyer
{attribute 'do_checks_for_implicit_code' := ''}
FUNCTION_BLOCK Unloading_Conveyer
VAR_OUTPUT
	/// TRUE sending a piece
	recv_O: BOOL;
	/// Spits out the data of the piece we just pulled
	Piece_Out: Piece;
END_VAR
VAR
	Found: BOOL;
	Target_Type: UINT;
	i: INT;
	j: INT;
END_VAR
VAR_INPUT
	/// Modbus index for the sensor
	Ioff: UINT;
	/// Modbus index for the motor
	Qoff: UINT;
	/// 1 = Top (W1), 2 = Bottom (W2)
	Target_WH: INT;
	/// 0 for going UP , 1 for going DOWN
	Direction: UINT;
	/// Command to fetch a piece
	Unload_Req: BOOL;
	///d TRUE if next belt empty~
	free_I: BOOL;
	piece_material: UINT;
	reg_numb: UINT;
END_VAR

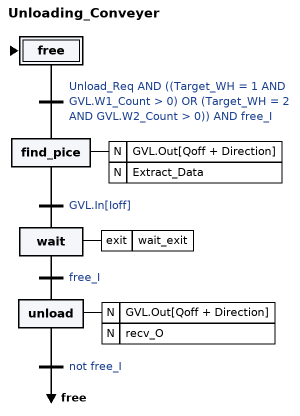
INITIAL_STEP free:
END_STEP
TRANSITION FROM free TO find_pice
    := Unload_Req AND ((Target_WH = 1 AND GVL.W1_Count > 0) OR (Target_WH = 2 AND GVL.W2_Count > 0)) AND free_I;
END_TRANSITION
STEP find_pice:
    GVL.Out[Qoff + Direction](N);
    Extract_Data(N);
END_STEP
TRANSITION FROM find_pice TO wait
    := GVL.In[Ioff];
END_TRANSITION
STEP wait:
    wait_exit(P0);  // exit action
END_STEP
TRANSITION FROM wait TO unload
    := free_I;
END_TRANSITION
STEP unload:
    GVL.Out[Qoff + Direction](N);
    recv_O(N);
END_STEP
TRANSITION FROM unload TO free
    := not free_I;
END_TRANSITION

ACTION Extract_Data:
IF NOT Found THEN
    Target_Type := piece_material;
    // --- TARGETING TOP WAREHOUSE (W1) ---
    IF Target_WH = 1 AND GVL.W1_Count > 0 THEN
        FOR i := 0 TO GVL.W1_Count - 1 DO
            IF Target_Type > 0 AND GVL.WareHouseTop[i].Type_ID = Target_Type THEN
                // Copy the piece data out to the conveyor belt
                Piece_Out := GVL.WareHouseTop[i];
                GVL.Reg[reg_numb] := GVL.WareHouseTop[i].Type_ID;
                // Shift remaining pieces to close the gap
                FOR j := i TO GVL.W1_Count - 2 DO
                    GVL.WareHouseTop[j] := GVL.WareHouseTop[j + 1];
                END_FOR;
                // Clear last slot
                GVL.WareHouseTop[GVL.W1_Count - 1].Type_ID := 0;
                GVL.WareHouseTop[GVL.W1_Count - 1].Is_Black := FALSE;
                // Update the counter and reset unload_type
                GVL.W1_Count := GVL.W1_Count - 1;
                piece_material := 0;
                Found := TRUE;
                EXIT;
            END_IF;
        END_FOR;
    // --- TARGETING BOTTOM WAREHOUSE (W2) ---
    ELSIF Target_WH = 2 AND GVL.W2_Count > 0 THEN
        FOR i := 0 TO GVL.W2_Count - 1 DO
            IF Target_Type > 0 AND GVL.WareHouseBottom[i].Type_ID = Target_Type THEN
                // Copy the piece data out to the conveyor belt
                Piece_Out := GVL.WareHouseBottom[i];
                GVL.Reg[reg_numb] := GVL.WareHouseBottom[i].Type_ID;
                // Shift remaining pieces to close the gap
                FOR j := i TO GVL.W2_Count - 2 DO
                    GVL.WareHouseBottom[j] := GVL.WareHouseBottom[j + 1];
                END_FOR;
                // Clear last slot
                GVL.WareHouseBottom[GVL.W2_Count - 1].Type_ID := 0;
                GVL.WareHouseBottom[GVL.W2_Count - 1].Is_Black := FALSE;
                // Update the counter and reset unload_type
                GVL.W2_Count := GVL.W2_Count - 1;
                piece_material := 0;
                Found := TRUE;
                EXIT;
            END_IF;
        END_FOR;
    END_IF;
END_IF;
END_ACTION

ACTION wait_exit:
GVL.Reg[reg_numb] := 0;
Found := FALSE;
END_ACTION

ACTION clear_vars:
GVL.Reg[reg_numb] := 0;
END_ACTION

END_FUNCTION_BLOCK

// Device/Application/Conveyers/Input_Conveyer
{attribute 'do_checks_for_implicit_code' := ''}
FUNCTION_BLOCK Input_Conveyer
VAR_OUTPUT
	/// TRUE when I have a piece at the end of my belt
	recv_O: BOOL;
	/// Spits out the data of the piece we just created
	Piece_Out: Piece;
END_VAR
VAR
	i: INT;
	v: INT;
END_VAR
VAR_INPUT
	/// Modbus index for the sensor at the drop zone
	Ioff: UINT;
	/// Modbus index for the motor 
	Qoff: UINT;
	/// Comand To Create Piece
	Create_Piece: BOOL;
	/// Piece Material
	piece_material: UINT;
	/// TRUE when next belt has no piece and can take one
	free_I: BOOL;
	/// Register number
	reg_numb: UINT;
END_VAR

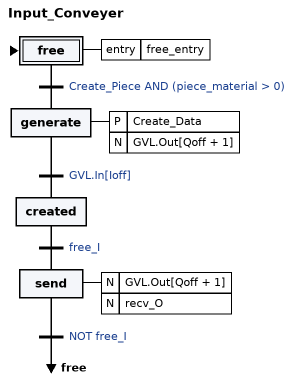
INITIAL_STEP free:
    free_entry(P1);  // entry action
END_STEP
TRANSITION FROM free TO generate
    := Create_Piece AND (piece_material > 0);
END_TRANSITION
STEP generate:
    Create_Data(P);
    GVL.Out[Qoff + 1](N);
END_STEP
TRANSITION FROM generate TO created
    := GVL.In[Ioff];
END_TRANSITION
STEP created:
END_STEP
TRANSITION FROM created TO send
    := free_I;
END_TRANSITION
STEP send:
    GVL.Out[Qoff + 1](N);
    recv_O(N);
END_STEP
TRANSITION FROM send TO free
    := NOT free_I;
END_TRANSITION

ACTION free_entry:
GVL.Reg[reg_numb] := 0;
Piece_Out.Type_ID := 0;
Piece_Out.Is_Black := FALSE;
END_ACTION

ACTION Create_Data:
// Generate the brand new piece data
GVL.Reg[reg_numb] := piece_material;
Piece_Out.Type_ID := piece_material;
Piece_Out.Is_Black := FALSE;
END_ACTION

END_FUNCTION_BLOCK

// Device/Application/Conveyers/Machine_Conveyer
{attribute 'do_checks_for_implicit_code' := ''}
FUNCTION_BLOCK Machine_Conveyer
VAR_OUTPUT
	Piece_Out: PIECE;
	free_O: BOOL;
	recv_O: BOOL;
END_VAR
VAR
	/// --- Memory for Assembly ---
	Saved_Top: UINT := 0;
	Saved_Leg1: UINT := 0;
	Saved_Leg2: UINT := 0;
	/// 0=Pass, 1=Transform, 2=Swallow, 3=Assemble
	Action_Type: UINT;
	Process_Time: TIME;
	Target_ID: UINT;
	/// Loop counter
	i: INT;
	/// --- Recipe Lookups ---
	Req_Top_ID: UINT;
	Req_Leg_ID: UINT;
	Req_Join_Tool: INT;
	/// Output: 0, 1, or 2 (Tells the 3D sim to rotate the tool)
	Needed_Tool: INT;
	/// True if the machine needs to change tools
	Needs_Rotation: BOOL;
	Active_Tool_Slot: INT := 0;
	Found: BOOL := TRUE;
	Working_Piece: Piece;
END_VAR
VAR_INPUT
	Ioff: UINT;
	Qoff: UINT;
	Piece_In: PIECE;
	recv_I: BOOL;
	free_I: BOOL;
	/// 0 for going UP , 1 for going DOWN
	Direction: UINT;
	/// e.g., [1, 2, 3]
	Tool_Magazine: ARRAY[0..2] OF INT;
END_VAR

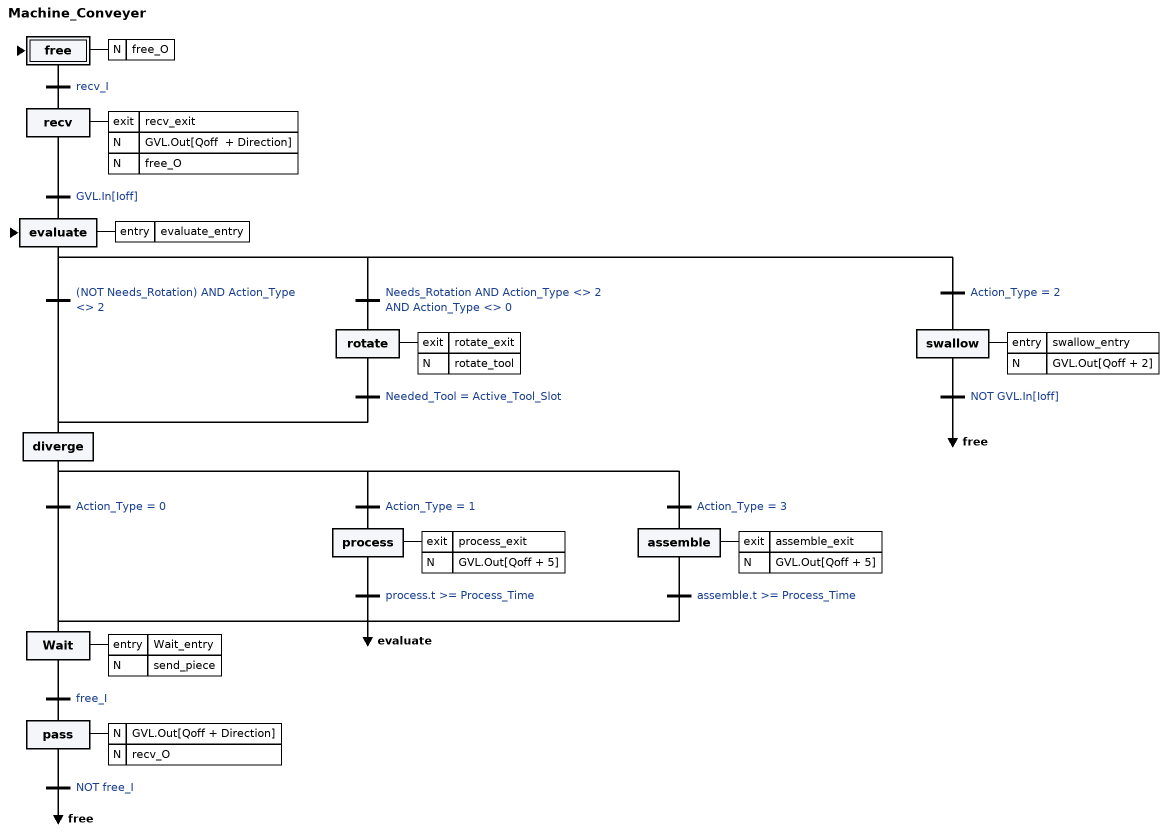
INITIAL_STEP free:
    free_O(N);
END_STEP
TRANSITION FROM free TO recv
    := recv_I;
END_TRANSITION
STEP recv:
    recv_exit(P0);  // exit action
    GVL.Out[Qoff  + Direction](N);
    free_O(N);
END_STEP
TRANSITION FROM recv TO evaluate
    := GVL.In[Ioff];
END_TRANSITION
STEP evaluate:
    evaluate_entry(P1);  // entry action
END_STEP
TRANSITION FROM evaluate TO diverge
    := (NOT Needs_Rotation) AND Action_Type <> 2;
END_TRANSITION
TRANSITION FROM evaluate TO rotate
    := Needs_Rotation AND Action_Type <> 2 AND Action_Type <> 0;
END_TRANSITION
STEP rotate:
    rotate_exit(P0);  // exit action
    rotate_tool(N);
END_STEP
TRANSITION FROM rotate TO diverge
    := Needed_Tool = Active_Tool_Slot;
END_TRANSITION
TRANSITION FROM evaluate TO swallow
    := Action_Type = 2;
END_TRANSITION
STEP swallow:
    swallow_entry(P1);  // entry action
    GVL.Out[Qoff + 2](N);
END_STEP
TRANSITION FROM swallow TO free
    := NOT GVL.In[Ioff];
END_TRANSITION
STEP diverge:
END_STEP
TRANSITION FROM diverge TO Wait
    := Action_Type = 0;
END_TRANSITION
TRANSITION FROM diverge TO process
    := Action_Type = 1;
END_TRANSITION
STEP process:
    process_exit(P0);  // exit action
    GVL.Out[Qoff + 5](N);
END_STEP
TRANSITION FROM process TO evaluate
    := process.t >= Process_Time;
END_TRANSITION
TRANSITION FROM diverge TO assemble
    := Action_Type = 3;
END_TRANSITION
STEP assemble:
    assemble_exit(P0);  // exit action
    GVL.Out[Qoff + 5](N);
END_STEP
TRANSITION FROM assemble TO Wait
    := assemble.t >= Process_Time;
END_TRANSITION
STEP Wait:
    Wait_entry(P1);  // entry action
    send_piece(N);
END_STEP
TRANSITION FROM Wait TO pass
    := free_I;
END_TRANSITION
STEP pass:
    GVL.Out[Qoff + Direction](N);
    recv_O(N);
END_STEP
TRANSITION FROM pass TO free
    := NOT free_I;
END_TRANSITION

ACTION send_piece:
Piece_Out := Working_Piece;
END_ACTION

ACTION recv_exit:
Working_Piece := Piece_In;
END_ACTION

ACTION Wait_entry:
Process_Time := GVL.Tool_Time[Tool_Magazine[Active_Tool_Slot]];
END_ACTION

ACTION update_creation_state:
// IF Action_Type = 1 THEN // We just finished a single transformation
//     IF Target_ID = 3 OR Target_ID = 4 OR Target_ID = 6 OR Target_ID = 7 THEN
//         GVL.Need_Top := FALSE; // Top is finished!
//     ELSIF Target_ID = 5 OR Target_ID = 8 THEN
//         GVL.Need_Legs := GVL.Need_Legs - 1; // One Leg is finished!
//     END_IF;
// END_IF;
END_ACTION

ACTION recv_entry:

END_ACTION

ACTION rotate_exit:
GVL.Out[Qoff + 3] := FALSE;
END_ACTION

ACTION evaluate_entry:
// // 1. Reset defaults
// Action_Type := 0; // Default: Pass it down the line
// Process_Time := T#0S;
// Target_ID := Working_Piece.Type_ID;
// 
// // 2. Decode the Global Target (What are we trying to build?)
// CASE GVL.Target_Table OF
//     9:  Req_Top_ID := 3; Req_Leg_ID := 5; Req_Join_Tool := 8; // RWW
//     10: Req_Top_ID := 4; Req_Leg_ID := 5; Req_Join_Tool := 8; // SWW
//     11: Req_Top_ID := 3; Req_Leg_ID := 8; Req_Join_Tool := 9; // RWM
//     12: Req_Top_ID := 4; Req_Leg_ID := 8; Req_Join_Tool := 9; // SWM
//     13: Req_Top_ID := 6; Req_Leg_ID := 8; Req_Join_Tool := 8; // RMM
//     14: Req_Top_ID := 7; Req_Leg_ID := 8; Req_Join_Tool := 8; // SMM
// END_CASE;
// 
// // ==============================================================
// // 3. ASSEMBLY CHECK: Can I swallow or join this piece?
// // ==============================================================
// FOR i := 0 TO 2 DO
//     IF Tool_Magazine[i] = Req_Join_Tool THEN // I have the right assembly tool!
// 
//         // If it's the Leg we need, and I need legs
//         IF Working_Piece.Type_ID = Req_Leg_ID THEN
//             IF Saved_Leg1 = 0 THEN
//                 Saved_Leg1 := Working_Piece.Type_ID; Needed_Tool := i; Action_Type := 2; // Swallow
//             ELSIF Saved_Leg2 = 0 THEN
//                 Saved_Leg2 := Working_Piece.Type_ID; Needed_Tool := i; Action_Type := 2; // Swallow
//             END_IF;
//         END_IF;
// 		
// 		// If it's the Top we need, and I don't have one yet
//         IF Working_Piece.Type_ID = Req_Top_ID AND Saved_Top = 0 THEN
//             Saved_Top := Working_Piece.Type_ID;
//             Needed_Tool := i;
//             Action_Type := 2; // Swallow it!
//         END_IF;
// 
//         // Do I have all 3 parts now?
//         IF Action_Type = 2 AND Saved_Top > 0 AND Saved_Leg1 > 0 AND Saved_Leg2 > 0 THEN
//             Action_Type := 3; // ASSEMBLE!
//             Process_Time := T#10S;
//             Target_ID := GVL.Target_Table; 
//         END_IF;
//         
//         IF Action_Type <> 0 THEN EXIT; END_IF; // Stop checking tools if we made a decision
//     END_IF;
// END_FOR;
// 
// // ==============================================================
// // 4. TRANSFORM CHECK: Can I create a missing piece?
// // ==============================================================
// // Only run this if we didn't just swallow the piece!
// IF Action_Type = 0 AND (Working_Piece.Type_ID = 1 OR Working_Piece.Type_ID = 2) THEN
//     
// FOR i := 0 TO 2 DO
//         
//         // PRIORITY 1: ALWAYS TRY TO MAKE THE LEGS FIRST!
//         IF GVL.Need_Legs > 0 THEN
//             IF (Working_Piece.Type_ID = 1 AND Req_Leg_ID = 5 AND Tool_Magazine[i] = 3) THEN // Make LegW (Fast)
//                 Needed_Tool := i; Process_Time := T#10S; Target_ID := 5; Action_Type := 1; EXIT;
//             ELSIF (Working_Piece.Type_ID = 1 AND Req_Leg_ID = 5 AND Tool_Magazine[i] = 10) THEN // Make LegW (Slow)
//                 Needed_Tool := i; Process_Time := T#30S; Target_ID := 5; Action_Type := 1; EXIT;
//             ELSIF (Working_Piece.Type_ID = 2 AND Req_Leg_ID = 8 AND Tool_Magazine[i] = 5) THEN // Make LegM (Fast)
//                 Needed_Tool := i; Process_Time := T#30S; Target_ID := 8; Action_Type := 1; EXIT;
//             ELSIF (Working_Piece.Type_ID = 2 AND Req_Leg_ID = 8 AND Tool_Magazine[i] = 11) THEN // Make LegM (Slow)
//                 Needed_Tool := i; Process_Time := T#40S; Target_ID := 8; Action_Type := 1; EXIT;
//             END_IF;
// 		// PRIORITY 2: ONLY MAKE THE TOP IF THE LEGS ARE DONE! (Need_Legs = 0)
//         ELSIF GVL.Need_Top AND GVL.Need_Legs = 0 AND Action_Type = 0 THEN
//             IF (Working_Piece.Type_ID = 1 AND Req_Top_ID = 3 AND Tool_Magazine[i] = 1) THEN // Make RTopW
//                 Needed_Tool := i; Process_Time := T#30S; Target_ID := 3; Action_Type := 1; EXIT;
//             ELSIF (Working_Piece.Type_ID = 1 AND Req_Top_ID = 4 AND Tool_Magazine[i] = 2) THEN // Make STopW
//                 Needed_Tool := i; Process_Time := T#20S; Target_ID := 4; Action_Type := 1; EXIT;
//             ELSIF (Working_Piece.Type_ID = 2 AND Req_Top_ID = 6 AND Tool_Magazine[i] = 4) THEN // Make RTopM
//                 Needed_Tool := i; Process_Time := T#35S; Target_ID := 6; Action_Type := 1; EXIT;
//             ELSIF (Working_Piece.Type_ID = 2 AND Req_Top_ID = 7 AND Tool_Magazine[i] = 6) THEN // Make STopM
//                 Needed_Tool := i; Process_Time := T#25S; Target_ID := 7; Action_Type := 1; EXIT;
//             END_IF;
//         END_IF;
//         
//     END_FOR;
// END_IF;
// 
// 
// Check if we need to physically rotate the tool before working
IF Action_Type = 1 OR Action_Type = 3 THEN
    IF Needed_Tool <> Active_Tool_Slot THEN
        Needs_Rotation := TRUE;
    ELSE
        Needs_Rotation := FALSE;
    END_IF;
ELSE
	Needs_Rotation := FALSE;
END_IF
END_ACTION

ACTION rotate_tool:

IF Needed_Tool <> Active_Tool_Slot THEN
	// 2. Watch the Tool Alignment Sensor (Ioff + 1)
	IF NOT GVL.In[Ioff + 1] THEN
		Found := FALSE;
	END_IF
	
	IF GVL.In[Ioff + 1] AND NOT Found THEN
		IF Active_Tool_Slot + 1 > 2 THEN
			Active_Tool_Slot := 0;
		ELSE
			Active_Tool_Slot := Active_Tool_Slot + 1;
		END_IF
		Found := TRUE;
	END_IF;
	
	// 1. Turn on the rotation motor
	GVL.Out[Qoff + 3] := TRUE;
END_IF
END_ACTION

ACTION process_exit:
// Officially transform the piece to its new ID!
Working_Piece.Type_ID := Target_ID;

// Tell the rest of the factory (GVL) that this piece is done!
// IF Target_ID = 3 OR Target_ID = 4 OR Target_ID = 6 OR Target_ID = 7 THEN
//     GVL.Need_Top := FALSE;              // The Top is ready!
// ELSIF Target_ID = 5 OR Target_ID = 8 THEN
//     GVL.Need_Legs := GVL.Need_Legs - 1; // One Leg is ready!
// END_IF;

Action_Type := 0;
END_ACTION

ACTION assemble_exit:
// 1. Officially transform the piece to its new ID!
Working_Piece.Type_ID := Target_ID;
Action_Type := 0;
Saved_Leg1 := 0;
Saved_Leg2 := 0;
END_ACTION

ACTION swallow_entry:
IF Saved_Leg1 = 0 THEN
    Saved_Leg1 := Working_Piece.Type_ID;
ELSIF Saved_Leg2 = 0 THEN
    Saved_Leg2 := Working_Piece.Type_ID;
END_IF;
END_ACTION

END_FUNCTION_BLOCK

// Device/Application/Conveyers/Linear_Conveyor
{attribute 'do_checks_for_implicit_code' := ''}
FUNCTION_BLOCK Linear_Conveyor
VAR_OUTPUT
	/// TRUE when this belt has no piece and can take one
	free_O: BOOL;
	/// TRUE when I have a piece at the end of my belt
	recv_O: BOOL;
	/// You need this to hand the data over to the next conveyor
	Passed_Piece: Piece;
END_VAR
VAR_INPUT
	/// Modbus index for the physical sensor on this conveyor
	Ioff: UINT;
	/// Modbus index for the physical motor on this conveyor
	Qoff: UINT;
	/// 0 for going UP , 1 for going DOWN
	Direction: UINT;
	/// The data of the piece coming in from the previous conveyor
	Piece_Type: Piece;
	/// TRUE when previus belt wants to send a piece
	recv_I: BOOL;
	/// TRUE when next belt has no piece and can take one
	free_I: BOOL;
END_VAR

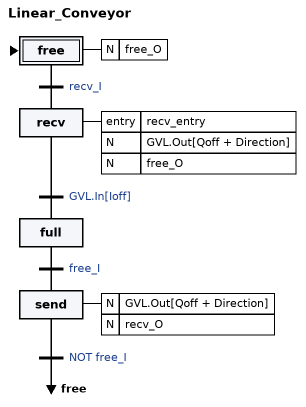
INITIAL_STEP free:
    free_O(N);
END_STEP
TRANSITION FROM free TO recv
    := recv_I;
END_TRANSITION
STEP recv:
    recv_entry(P1);  // entry action
    GVL.Out[Qoff + Direction](N);
    free_O(N);
END_STEP
TRANSITION FROM recv TO full
    := GVL.In[Ioff];
END_TRANSITION
STEP full:
END_STEP
TRANSITION FROM full TO send
    := free_I;
END_TRANSITION
STEP send:
    GVL.Out[Qoff + Direction](N);
    recv_O(N);
END_STEP
TRANSITION FROM send TO free
    := NOT free_I;
END_TRANSITION

ACTION recv_entry:
Passed_Piece := Piece_Type;
END_ACTION

END_FUNCTION_BLOCK

// Device/Application/SCADA_PRG
PROGRAM SCADA_PRG
VAR
    eActiveMode      : INT := 0;
    eCurrentTool     : INT := 1;
    eRequestedTool   : INT := 0;
    tonToolChange    : TON;
    bToolChangeBusy  : BOOL;
    tonIdleAlarm     : TON;
    bProcessingDone  : BOOL;
    old_Auto     : BOOL;
    old_Manual   : BOOL;
    old_Maint    : BOOL;
    old_T1       : BOOL;
    old_T2       : BOOL;
    old_T3       : BOOL;
    old_Done     : BOOL;
    old_Sensor   : BOOL;
END_VAR

(* === 1. MIRROR GVL I/O -> MODBUS COILS === *)
In_on         := GVL.Out[28];
M1a_on        := GVL.Out[70];
L1_on         := GVL.Out[80];
M1b_on        := GVL.Out[82];
L2_on         := GVL.Out[92];
M1c_on        := GVL.Out[94];
Out_on        := GVL.Out[48];

C1_In_Sensor  := GVL.In[11];
M1a_Sensor    := GVL.In[30];
C1_L1_Sensor  := GVL.In[36];
M1b_Sensor    := GVL.In[37];
C1_L2_Sensor  := GVL.In[43];
M1c_Sensor    := GVL.In[44];
C1_Out_Sensor := GVL.In[44];

(* === 2. OPERATING MODE INTERLOCKING === *)
IF M1a_Auto AND NOT old_Auto THEN
    eActiveMode := 1; M1a_Auto := FALSE;
END_IF
IF M1a_Manual AND NOT old_Manual THEN
    eActiveMode := 2; M1a_Manual := FALSE;
END_IF
IF M1a_Manutencao AND NOT old_Maint THEN
    eActiveMode := 3; M1a_Manutencao := FALSE;
END_IF

old_Auto   := M1a_Auto;
old_Manual := M1a_Manual;
old_Maint  := M1a_Manutencao;

(* === 3. TOOL CHANGE (Manual mode, 30s) === *)
IF M1a_T1 AND NOT old_T1 AND eActiveMode = 2 AND NOT bToolChangeBusy THEN
    eRequestedTool := 1; M1a_T1 := FALSE;
END_IF
IF M1a_T2 AND NOT old_T2 AND eActiveMode = 2 AND NOT bToolChangeBusy THEN
    eRequestedTool := 2; M1a_T2 := FALSE;
END_IF
IF M1a_T3 AND NOT old_T3 AND eActiveMode = 2 AND NOT bToolChangeBusy THEN
    eRequestedTool := 3; M1a_T3 := FALSE;
END_IF

old_T1 := M1a_T1;
old_T2 := M1a_T2;
old_T3 := M1a_T3;

IF eRequestedTool > 0 AND eRequestedTool <> eCurrentTool AND NOT bToolChangeBusy THEN
    bToolChangeBusy := TRUE;
END_IF

tonToolChange(IN := bToolChangeBusy, PT := T#30S);
IF tonToolChange.Q THEN
    eCurrentTool   := eRequestedTool;
    eRequestedTool := 0;
    bToolChangeBusy := FALSE;
END_IF

M1a_T1 := (eCurrentTool = 1);
M1a_T2 := (eCurrentTool = 2);
M1a_T3 := (eCurrentTool = 3);

(* === 4. MANUAL OPERATION DONE === *)
IF M1a_done AND NOT old_Done THEN
    bProcessingDone := TRUE; M1a_done := FALSE;
END_IF
old_Done := M1a_done;

IF old_Sensor AND NOT M1a_Sensor THEN
    bProcessingDone := FALSE;
END_IF
old_Sensor := M1a_Sensor;

(* === 5. IDLE ALARM (10s) === *)
tonIdleAlarm(IN := M1a_Sensor AND bProcessingDone, PT := T#10S);
M1a_Idle_Alarm := tonIdleAlarm.Q;

END_PROGRAM

// Device/Application/PRG_MQTT
PROGRAM PRG_MQTT
VAR
END_VAR

(*
  PRG_MQTT — MQTT telemetry publisher and RPC subscriber
  Paste into the IMPLEMENTATION (lower) section of PRG_MQTT.
  Call PRG_MQTT from MainTask once per scan.

  One publish group is sent every 500ms. Four groups cycle every 2s.
  The FB is called ONCE per scan so R_TRIG fires correctly each time.
*)

// ── Publisher configuration ───────────────────────────────────────────────
GVL_MQTT.fbMQTT_Pub.i_xEnable        := TRUE;
GVL_MQTT.fbMQTT_Pub.i_sBrokerAddress := 'thingsboard.cloud';
GVL_MQTT.fbMQTT_Pub.i_uiPort         := 1883;
GVL_MQTT.fbMQTT_Pub.i_sUsername      := 'lv33yCUTuUp9BiERh8bJ';
GVL_MQTT.fbMQTT_Pub.i_sPassword      := '';
GVL_MQTT.fbMQTT_Pub.i_sClientID      := 'codesys-plc-pub';
GVL_MQTT.fbMQTT_Pub.i_sTopicPublish  := 'v1/devices/me/telemetry';
GVL_MQTT.fbMQTT_Pub.i_xRetain        := FALSE;
GVL_MQTT.fbMQTT_Pub.i_xAutoReconnect := TRUE;

// ── Subscriber configuration ──────────────────────────────────────────────
GVL_MQTT.fbMQTT_Sub.i_xEnable         := TRUE;
GVL_MQTT.fbMQTT_Sub.i_sBrokerAddress  := 'thingsboard.cloud';
GVL_MQTT.fbMQTT_Sub.i_uiPort          := 1883;
GVL_MQTT.fbMQTT_Sub.i_sUsername       := 'YN1hLdTh20UMCIGUIhTQ';
GVL_MQTT.fbMQTT_Sub.i_sPassword       := '';
GVL_MQTT.fbMQTT_Sub.i_sClientID       := 'codesys-plc-sub';
GVL_MQTT.fbMQTT_Sub.i_sTopicSubscribe := 'v1/devices/me/rpc/request/+';
GVL_MQTT.fbMQTT_Sub.i_xSubscribe      := TRUE;
GVL_MQTT.fbMQTT_Sub.i_xAutoReconnect  := TRUE;

// ── Advance to next group every 500ms ────────────────────────────────────
GVL_MQTT.tPublishTimer(IN := TRUE, PT := T#500MS);

IF GVL_MQTT.tPublishTimer.Q THEN
    GVL_MQTT.tPublishTimer(IN := FALSE);

    GVL_MQTT.nPublishGroup := GVL_MQTT.nPublishGroup + 1;
    IF GVL_MQTT.nPublishGroup > 4 THEN
        GVL_MQTT.nPublishGroup := 1;
    END_IF

    CASE GVL_MQTT.nPublishGroup OF

    1: // Input line signals
        MQTT_Client.FC_AddKeyValueToJSON(i_sKeyToAdd := 'create_piece_I1',   i_sValueToAdd := BOOL_TO_STRING(PLC_PRG.Create_Piece_I1));
        MQTT_Client.FC_AddKeyValueToJSON(i_sKeyToAdd := 'create_piece_I2',   i_sValueToAdd := BOOL_TO_STRING(PLC_PRG.Create_Piece_I2));
        MQTT_Client.FC_AddKeyValueToJSON(i_sKeyToAdd := 'create_piece_I3',   i_sValueToAdd := BOOL_TO_STRING(PLC_PRG.Create_Piece_I3));
        MQTT_Client.FC_AddKeyValueToJSON(i_sKeyToAdd := 'create_piece_I4',   i_sValueToAdd := BOOL_TO_STRING(PLC_PRG.Create_Piece_I4));
        MQTT_Client.FC_AddKeyValueToJSON(i_sKeyToAdd := 'piece_material_I1', i_sValueToAdd := WORD_TO_STRING(PLC_PRG.piece_material_I1));
        MQTT_Client.FC_AddKeyValueToJSON(i_sKeyToAdd := 'piece_material_I2', i_sValueToAdd := WORD_TO_STRING(PLC_PRG.piece_material_I2));
        MQTT_Client.FC_AddKeyValueToJSON(i_sKeyToAdd := 'piece_material_I3', i_sValueToAdd := WORD_TO_STRING(PLC_PRG.piece_material_I3));
        MQTT_Client.FC_AddKeyValueToJSON(i_sKeyToAdd := 'piece_material_I4', i_sValueToAdd := WORD_TO_STRING(PLC_PRG.piece_material_I4));
        GVL_MQTT.fbMQTT_Pub.i_sPayload := MQTT_Client.FC_CreateJSON();
        GVL_MQTT.fbMQTT_Pub.i_xPublish := TRUE;

    2: // Unload request signals
        MQTT_Client.FC_AddKeyValueToJSON(i_sKeyToAdd := 'unload_req_U1',  i_sValueToAdd := BOOL_TO_STRING(PLC_PRG.Unload_Req_U1));
        MQTT_Client.FC_AddKeyValueToJSON(i_sKeyToAdd := 'unload_req_U2',  i_sValueToAdd := BOOL_TO_STRING(PLC_PRG.Unload_Req_U2));
        MQTT_Client.FC_AddKeyValueToJSON(i_sKeyToAdd := 'unload_req_U3',  i_sValueToAdd := BOOL_TO_STRING(PLC_PRG.Unload_Req_U3));
        MQTT_Client.FC_AddKeyValueToJSON(i_sKeyToAdd := 'unload_req_U4',  i_sValueToAdd := BOOL_TO_STRING(PLC_PRG.Unload_Req_U4));
        MQTT_Client.FC_AddKeyValueToJSON(i_sKeyToAdd := 'unload_req_U5',  i_sValueToAdd := BOOL_TO_STRING(PLC_PRG.Unload_Req_U5));
        MQTT_Client.FC_AddKeyValueToJSON(i_sKeyToAdd := 'unload_req_U6',  i_sValueToAdd := BOOL_TO_STRING(PLC_PRG.Unload_Req_U6));
        MQTT_Client.FC_AddKeyValueToJSON(i_sKeyToAdd := 'unload_req_U7',  i_sValueToAdd := BOOL_TO_STRING(PLC_PRG.Unload_Req_U7));
        MQTT_Client.FC_AddKeyValueToJSON(i_sKeyToAdd := 'unload_req_U8',  i_sValueToAdd := BOOL_TO_STRING(PLC_PRG.Unload_Req_U8));
        MQTT_Client.FC_AddKeyValueToJSON(i_sKeyToAdd := 'unload_req_U9',  i_sValueToAdd := BOOL_TO_STRING(PLC_PRG.Unload_Req_U9));
        MQTT_Client.FC_AddKeyValueToJSON(i_sKeyToAdd := 'unload_req_U10', i_sValueToAdd := BOOL_TO_STRING(PLC_PRG.Unload_Req_U10));
        GVL_MQTT.fbMQTT_Pub.i_sPayload := MQTT_Client.FC_CreateJSON();
        GVL_MQTT.fbMQTT_Pub.i_xPublish := TRUE;

    3: // Unload material type per dock
        MQTT_Client.FC_AddKeyValueToJSON(i_sKeyToAdd := 'unload_type_U1',  i_sValueToAdd := WORD_TO_STRING(PLC_PRG.Unload_Type_U1));
        MQTT_Client.FC_AddKeyValueToJSON(i_sKeyToAdd := 'unload_type_U2',  i_sValueToAdd := WORD_TO_STRING(PLC_PRG.Unload_Type_U2));
        MQTT_Client.FC_AddKeyValueToJSON(i_sKeyToAdd := 'unload_type_U3',  i_sValueToAdd := WORD_TO_STRING(PLC_PRG.Unload_Type_U3));
        MQTT_Client.FC_AddKeyValueToJSON(i_sKeyToAdd := 'unload_type_U4',  i_sValueToAdd := WORD_TO_STRING(PLC_PRG.Unload_Type_U4));
        MQTT_Client.FC_AddKeyValueToJSON(i_sKeyToAdd := 'unload_type_U5',  i_sValueToAdd := WORD_TO_STRING(PLC_PRG.Unload_Type_U5));
        MQTT_Client.FC_AddKeyValueToJSON(i_sKeyToAdd := 'unload_type_U6',  i_sValueToAdd := WORD_TO_STRING(PLC_PRG.Unload_Type_U6));
        MQTT_Client.FC_AddKeyValueToJSON(i_sKeyToAdd := 'unload_type_U7',  i_sValueToAdd := WORD_TO_STRING(PLC_PRG.Unload_Type_U7));
        MQTT_Client.FC_AddKeyValueToJSON(i_sKeyToAdd := 'unload_type_U8',  i_sValueToAdd := WORD_TO_STRING(PLC_PRG.Unload_Type_U8));
        MQTT_Client.FC_AddKeyValueToJSON(i_sKeyToAdd := 'unload_type_U9',  i_sValueToAdd := WORD_TO_STRING(PLC_PRG.Unload_Type_U9));
        MQTT_Client.FC_AddKeyValueToJSON(i_sKeyToAdd := 'unload_type_U10', i_sValueToAdd := WORD_TO_STRING(PLC_PRG.Unload_Type_U10));
        GVL_MQTT.fbMQTT_Pub.i_sPayload := MQTT_Client.FC_CreateJSON();
        GVL_MQTT.fbMQTT_Pub.i_xPublish := TRUE;

    4: // Warehouse counts
        MQTT_Client.FC_AddKeyValueToJSON(i_sKeyToAdd := 'W1_count', i_sValueToAdd := WORD_TO_STRING(GVL.W1_Count));
        MQTT_Client.FC_AddKeyValueToJSON(i_sKeyToAdd := 'W2_count', i_sValueToAdd := WORD_TO_STRING(GVL.W2_Count));
        GVL_MQTT.fbMQTT_Pub.i_sPayload := MQTT_Client.FC_CreateJSON();
        GVL_MQTT.fbMQTT_Pub.i_xPublish := TRUE;

    END_CASE
END_IF

// ── Call publisher FB once per scan ──────────────────────────────────────
GVL_MQTT.fbMQTT_Pub();

// Drop publish trigger after one scan so R_TRIG resets correctly
IF GVL_MQTT.fbMQTT_Pub.i_xPublish THEN
    GVL_MQTT.fbMQTT_Pub.i_xPublish := FALSE;
END_IF

// ── Call subscriber FB once per scan ─────────────────────────────────────
GVL_MQTT.fbMQTT_Sub();

// ── Handle incoming RPC commands ─────────────────────────────────────────
IF GVL_MQTT.fbMQTT_Sub.q_xReceivedMessageNotification THEN
    GVL_MQTT.sRPCMessage := GVL_MQTT.fbMQTT_Sub.q_sLastReceivedMessage;
    GVL_MQTT.bNewRPC     := TRUE;
END_IF

END_PROGRAM

// Device/Application/AlarmManager
PROGRAM AlarmManager

// ── M1a Idle Workpiece Alarm ──
// GVL.TON_M1a(IN := GVL.M1a_done AND GVL.Out[8], PT := T#10S);
// GVL.M1a_Idle_Alarm := GVL.TON_M1a.Q;

// ── M1b Idle Workpiece Alarm ──
// GVL.TON_M1b(IN := GVL.M1b_done AND GVL.Out[10], PT := T#10S);
// GVL.M1b_Idle_Alarm := GVL.TON_M1b.Q;

// ── M1c Idle Workpiece Alarm ──
// GVL.TON_M1c(IN := GVL.M1c_done AND GVL.Out[12], PT := T#10S);
// GVL.M1c_Idle_Alarm := GVL.TON_M1c.Q;


// ── Write alarm outputs into Modbus Out[] buffer ──
// GVL.Out[215] := GVL.M1a_done;
// GVL.Out[216] := GVL.M1b_done;
// GVL.Out[217] := GVL.M1c_done;
// GVL.Out[218] := GVL.M1a_Idle_Alarm;
// GVL.Out[219] := GVL.M1b_Idle_Alarm;
// GVL.Out[220] := GVL.M1c_Idle_Alarm;

END_PROGRAM
